(* IEC 61131-3 sources: PortalRobot/Portal_robot/Device/application/FB/FB_CELL_MANAGER, 14 files *)

(* ---- FB_CELL_MANAGER.st ---- *)
FUNCTION_BLOCK FB_CELL_MANAGER
VAR_INPUT
	xIoManual : BOOL; // Прямой ручной слой отменяет задание, не сбрасывая аварии
	axMagazineAutoSwapPending : ARRAY [1..GVL_CELL_SETTINGS.MagazineCount] OF BOOL; // Палета ждёт окна обмена
	axMagazineExchangeInProgress : ARRAY [1..GVL_CELL_SETTINGS.MagazineCount] OF BOOL; // Во время смены палет запрещены операции только с этим магазином
	xMagazineExchangeActive : BOOL; // Есть активный обмен палет; подавляет временные предупреждения о запасах
	xStart            : BOOL; // Импульс запуска цикла или отмены остановки
	xStop             : BOOL; // Импульс контролируемой остановки
	xTestAbort        : BOOL; // Немедленная отмена только тестового прогона
	xResetRequest     : BOOL; // Необработанный запрос сброса от HMI
	xReset            : BOOL; // Общий сброс владельцев ошибок
	xOperatorChoice   : BOOL; // Импульс ответа активному предпусковому опросу
	xOperatorCancel   : BOOL; // Импульс отмены предпускового опроса
	uiOperatorChoice  : UINT; // Выбранное содержимое, тип продукции или станок
	xManual           : BOOL; // Ручной режим ячейки
	xIoDoRejected : BOOL;
    xIoEmergencyResetRejected : BOOL;
    xIoEmergencyStopActive : BOOL;
	xIoOverrideRejected : BOOL; // Отклонённая транзакция диагностики, эффект WARNING
	xSettingsRejected : BOOL; // Rejected or expired setting transaction
	uiModeRejectReason : UINT; // Одноцикловый отказ транзакции режима: 2 цикл, 3 Safety
	xGlobalError      : BOOL; // Глобальная ошибка ячейки
	xSafetyReady      : BOOL; // Все дискретные условия безопасности выполнены
	xDrivesReady      : BOOL; // Приводы готовы
	xMotionBusy       : BOOL; // Оси ещё движутся
	xRobotInterfaceReady : BOOL; // Выбранный интерфейс робота готов к работе
	lrRobotActualX    : LREAL; // Фактическая координата робота X
	lrRobotActualY    : LREAL; // Фактическая координата робота Y
	lrRobotActualZ    : LREAL; // Фактическая координата робота Z
	stSafetyHomePoint : ST_POINT; // Настроенная безопасная точка повторного запуска
	lrSafetyHomeToleranceX : LREAL; // Допуск HOME_SAFETY по X
	lrSafetyHomeToleranceY : LREAL; // Допуск HOME_SAFETY по Y
	lrSafetyHomeToleranceZ : LREAL; // Допуск HOME_SAFETY по Z
	lrStoppedPoseTolerance : LREAL; // Допуск контроля позы после штатной остановки
	Config            : ST_MULTI_TYPE_CONFIG; // Активная конфигурация типов
	xConfigurationValid : BOOL; // Конфигурация типов прошла проверку
	xPointsConfigured : BOOL; // HOME_SAFETY и точки включённого оборудования настроены
	stRobotStatus     : ST_ROBOT_STATUS; // Состояние робота
	astMagazineStatus : ARRAY [1..GVL_CELL_SETTINGS.MagazineCount] OF ST_MAGAZINE_STATUS;
	astMachineStatus  : ARRAY [1..3] OF ST_MACHINE_PUBLIC; // Состояния станков
	astMachineDiag    : ARRAY [1..3] OF ST_MACHINE_DIAG; // Автоматы станков
	FaultRequest      : ST_CELL_FAULT_REQUEST; // Диагностическая инъекция
END_VAR
VAR_OUTPUT
	Command            : ST_CELL_COMMAND; // Команды существующим блокам ячейки
	Status             : ST_CELL_STATUS; // Общий контракт состояния ячейки
	Diag               : ST_CELL_DIAG; // Общий контракт диагностики ячейки
	Error              : ST_CELL_ERRORS; // Общий контракт ошибок ячейки
	CycleStatus        : ST_CELL_CYCLE_STATUS; // Расширенная диагностика универсального цикла
	FaultStatus        : ST_FAULT_INJECTION_STATUS; // Инъекция логической ошибки ячейки
	uiReturnMagazine   : UINT; // Внутренний владелец парного цикла до возврата детали; 0 — цикл освобождён
END_VAR
VAR
	axGeometryUnloadBlocked : ARRAY [1..3] OF BOOL; // Вызванная деталь ждёт доступного свободного ГК
	atonGeometryWait : ARRAY [1..3] OF TON;
	audiGeometryWaitCallId : ARRAY [1..3] OF UDINT;
	axGeometryWaitWarned : ARRAY [1..3] OF BOOL;
	xGeometryHeld : BOOL;
	xGeometryDetailCounted : BOOL;
	uiGeometryMachine : UINT;
	uiGeometryStation : UINT;
	uiGeometryParkStation : UINT;
	uiGeometryStep : UINT;
	uiGeometryBypassReason : UINT;
	uiGeometryIndex : UINT;
	udiGeometryMagazineCounter : UDINT;
	eGeometryReturnState : E_CELL_MANAGER_STATE;
	eGeometrySafePoint : E_POINT_NAME;
	eGeometryChangePoint : E_POINT_NAME;
	eGeometryPlacePoint : E_POINT_NAME;
	xActiveMagazineAutoSwapPending : BOOL; // Удержать владельца и цикл до обмена его палеты
	eState               : E_CELL_MANAGER_STATE := E_CELL_MANAGER_STATE.IDLE; // Состояние универсального автомата
	eMagazineOperation   : E_MAGAZINE_OPERATION; // Выполняемая операция магазина
	eMachineOperation    : E_MACHINE_OPERATION; // Зафиксированная операция станка
	xRunning             : BOOL; // Защёлка автоматического цикла
	xStopRequested       : BOOL; // Остановка после безопасного шага
	xReadyToStart        : BOOL; // Условия запуска выполнены
	xRobotReady          : BOOL; // Робот готов принять маршрут
	xMagazineReady       : BOOL; // Магазин готов к операции
	xActiveMagazineExchangeInProgress : BOOL; // Выбранный магазин сейчас меняет палеты
	stMagazineStatus     : ST_MAGAZINE_STATUS; // Снимок выбранного магазина для существующего автомата
	uiActiveMagazine     : UINT; // Магазин текущей команды роботу
	uiSupplyMagazine     : UINT; // Источник следующих заготовок сохраняется между парными циклами
	xMagazine1Available  : BOOL;
	xMagazine2Available  : BOOL;
	xMagazineSelectionAllowed : BOOL; // Новое владение допускается только между операциями
	xMagazine1CanContinue : BOOL; // Первый магазин позволяет следующий технологический шаг
	xMagazine2CanContinue : BOOL; // Второй магазин позволяет следующий технологический шаг
	xMagazine1CanSupplyBlank : BOOL; // М1 позволяет штатный план TAKE перед отдельной выгрузкой
	xMagazine2CanSupplyBlank : BOOL; // М2 позволяет штатный план TAKE перед отдельной выгрузкой
	xMagazine1CanExchangeDetail : BOOL; // Заготовка М1 освобождает слот для детали робота
	xMagazine2CanExchangeDetail : BOOL;
	xMagazine1CanPutDetail : BOOL; // Готовый магазин со свободным местом для детали робота
	xMagazine2CanPutDetail : BOOL;
	xActiveMagazineCanExchangeDetail : BOOL;
	xHeldBlankLoadAvailable : BOOL; // При двух грузах можно сначала загрузить пустой станок
	uiMagazineType       : UINT; // Тип станка при проверке содержимого обоих магазинов
	uiPreferredMagazine  : UINT; // Назначение с учётом владельца цикла и сохранённого источника
	xReselectMagazine    : BOOL; // Требуется передать владение подходящему магазину
	xAlternateMagazineAvailable : BOOL; // Второй магазин готов принять непрерывный автоматический цикл
	xUseAlternateMagazineForDetail : BOOL; // У текущего магазина нет слота детали, у второго есть
	xAnyMagazineDetailSlotAvailable : BOOL; // Есть доступный слот детали хотя бы в одном магазине
	xNoDetailDestinationCondition : BOOL; // Робот держит готовую деталь без доступного слота
	xNoBlankStockCondition : BOOL; // Нет заготовок и текущей работы для автоматического цикла
	xDetailDestinationWarningActive : BOOL; // Предупреждение об отсутствии места уже выдано
	xBlankStockWarningActive : BOOL; // Предупреждение об отсутствии заготовок уже выдано
	xMachineWorkPending : BOOL; // Станок занят/обрабатывает, запускается или содержит изделие
	xAnyMachineBusy      : BOOL; // Хотя бы один станок обслуживается
	xMachineServiceStarted : BOOL; // Выбранный станок вошёл в рецепт
	xReselectAfterRobotRelease : BOOL; // После снятия команды требуется повторный выбор
	xChangePrepared      : BOOL; // Для CHANGE зафиксированы совместимый станок и два корректных слота
	xFaultAllowed        : BOOL; // Инъекция разрешена в полностью остановленной ячейке
	xResetAllowed        : BOOL; // Локальная ошибка может быть сброшена
	xPayloadRouteWarningActive : BOOL; // Предупреждение о несовпадении типа груза и назначения уже выдано
	xPrestartGripper1Occupied : BOOL; // Снимок занятости первого захвата на момент запуска опроса
	xPrestartGripper2Occupied : BOOL; // Снимок занятости второго захвата на момент запуска опроса
	xSafetyHomeRequired : BOOL; // Защёлка обязательного возврата в HOME_SAFETY
	xRobotAtSafetyHome  : BOOL; // Робот находится в допустимом диапазоне HOME_SAFETY
	xStoppedPoseValid   : BOOL; // После штатной остановки сохранена доверенная поза
	xWasRunning         : BOOL; // Состояние цикла на предыдущем вызове
	xStartCheckCellIdle           : BOOL; // Отдельные условия запуска для HMI
	xStartCheckAutomaticMode      : BOOL;
	xStartCheckNoBlockingError    : BOOL;
	xStartCheckRobotInterfaceReady: BOOL;
	xStartCheckConfigurationValid : BOOL;
	xStartCheckPointsConfigured   : BOOL;
	xStartCheckDrivesReady        : BOOL;
	xStartCheckRobotReady         : BOOL;
	xStartCheckMagazineReady      : BOOL;
	xStartCheckTaskAvailable      : BOOL;
	xStartCheckSafetyHome         : BOOL;
	xStartCheckSafety             : BOOL;
	xOperatorPromptState          : BOOL; // Текущий шаг ожидает ответ HMI
	xOperatorChoiceAllowed        : BOOL;
	xOperatorCancelAllowed        : BOOL;
	uiOperatorPrompt              : UINT;
	uiOperatorTypeMask            : UINT;
	uiOperatorMachineMask         : UINT;
	uiStartConditionsMet         : UINT;
	lrStoppedPoseX      : LREAL; // Доверенная координата X штатной остановки
	lrStoppedPoseY      : LREAL; // Доверенная координата Y штатной остановки
	lrStoppedPoseZ      : LREAL; // Доверенная координата Z штатной остановки
	uiReadyMachines      : UINT; // Число доступных маршрутных целей
	uiMachine            : UINT; // Индекс станка
	uiMagazineIndex      : UINT; // Индекс магазина при поиске свободного слота
	uiCandidateMachine   : UINT; // Результат выбора
	uiSelectedMachine    : UINT; // Зафиксированный станок
	uiSelectedType       : UINT; // Тип маршрута
	uiBlankPayloadType   : UINT; // Тип заготовки в первом захвате
	uiDetailPayloadType  : UINT; // Тип готовой детали во втором захвате
	axMachineStartPending: ARRAY [1..3] OF BOOL; // Станок обслужен, но xProcessing ещё не подтверждён
	iTakeSlot            : SINT; // Зарезервированный слот заготовки
	iPutSlot             : SINT; // Зарезервированный слот укладки
	iTakeOriginSlot      : SINT; // Исходный слот заготовки для приоритетного возврата
	rtStart              : R_TRIG; // Фронт запуска
	rtStop               : R_TRIG; // Фронт остановки
	rtReset              : R_TRIG; // Фронт сброса
	rtOperatorChoice     : R_TRIG; // Один ответ не переносится на следующий шаг опроса
	rtOperatorCancel     : R_TRIG; // Фронт отмены предпускового опроса
	fbFaultInjector      : FB_CELL_FAULT_INJECTOR; // Проверка противоречивого груза
END_VAR
VAR CONSTANT
	FIRST_MACHINE     : UINT := UINT#1;
	LAST_MACHINE      : UINT := UINT#3;
	MACHINE_SWITCH_DEADBAND : TIME := T#1S; // Минимальный выигрыш времени для смены ожидаемой цели
	START_PENDING_ESTIMATE  : TIME := T#1S; // Оценка перехода от освобождения робота до xProcessing
	ERR_BOTH_GRIPPERS : DWORD := DWORD#16#0000_0001;
	ERR_ROBOT         : DWORD := DWORD#16#0000_0002;
	ERR_MAGAZINE      : DWORD := DWORD#16#0000_0004;
	ERR_MACHINE       : DWORD := DWORD#16#0000_0008;
	ERR_GLOBAL_STOP   : DWORD := DWORD#16#0000_0010;
	WRN_START_NOT_READY       : UINT := UINT#4;
	WRN_STOP_NOT_RUNNING      : UINT := UINT#5;
	WRN_SIM_ERROR_NOT_ALLOWED : UINT := UINT#8;
	WRN_PAYLOAD_ROUTE_MISMATCH : UINT := UINT#9;
	WRN_SAFETY_HOME_REQUIRED   : UINT := UINT#10;
	WRN_MANUAL_MODE_REJECTED   : UINT := UINT#11;
	WRN_CELL_SETTING_REJECTED : UINT := UINT#28;
	WRN_AUTOMATIC_MODE_REJECTED : UINT := UINT#27; // WARNING: общая авария удерживает ручной режим
	WRN_GRIPPER1_CONTENT       : UINT := UINT#15;
	WRN_GRIPPER2_CONTENT       : UINT := UINT#16;
	WRN_PAYLOAD_TYPE_CHOICE    : UINT := UINT#17;
	WRN_DETAIL_SLOT_REQUIRED   : UINT := UINT#18;
	WRN_START_MACHINE_REQUIRED : UINT := UINT#19;
	WRN_START_MACHINE_CHOICE   : UINT := UINT#20;
	WRN_OPERATOR_REPLY_REJECTED: UINT := UINT#21;
	WRN_OPERATOR_CANCEL_REJECTED: UINT := UINT#22;
	WRN_NO_DETAIL_DESTINATION  : UINT := UINT#29;
	WRN_NO_BLANK_STOCK         : UINT := UINT#30;
	WRN_GEOMETRY_WAIT_TIMEOUT  : UINT := UINT#52;
	WRN_IO_OVERRIDE_REJECTED   : UINT := UINT#31;
    WRN_IO_DO_REJECTED : UINT := UINT#32;
    WRN_IO_EMERGENCY_RESET_REJECTED : UINT := UINT#33;
END_VAR

// --- BEGIN IMPLEMENTATION ---

IF xIoDoRejected THEN
    Diag.stWarning.uiCode := WRN_IO_DO_REJECTED; // WARNING: вход/команда прямого ручного I/O не применены
    Diag.stWarning.udiSequence := Diag.stWarning.udiSequence + UDINT#1;
    IF Diag.stWarning.udiSequence = UDINT#0 THEN Diag.stWarning.udiSequence := UDINT#1; END_IF;
END_IF;
IF xIoEmergencyResetRejected THEN
    Diag.stWarning.uiCode := WRN_IO_EMERGENCY_RESET_REJECTED; // WARNING: останов остаётся
    Diag.stWarning.udiSequence := Diag.stWarning.udiSequence + UDINT#1;
    IF Diag.stWarning.udiSequence = UDINT#0 THEN Diag.stWarning.udiSequence := UDINT#1; END_IF;
END_IF;
IF xIoOverrideRejected THEN
    Diag.stWarning.uiCode := WRN_IO_OVERRIDE_REJECTED; // WARNING: входы не изменены
    Diag.stWarning.udiSequence := Diag.stWarning.udiSequence + UDINT#1;
    IF Diag.stWarning.udiSequence = UDINT#0 THEN Diag.stWarning.udiSequence := UDINT#1; END_IF;
END_IF;
IF xSettingsRejected THEN
	Diag.stWarning.uiCode := WRN_CELL_SETTING_REJECTED; // WARNING: settings unchanged
	Diag.stWarning.udiSequence := Diag.stWarning.udiSequence + UDINT#1;
	IF Diag.stWarning.udiSequence = UDINT#0 THEN Diag.stWarning.udiSequence := UDINT#1; END_IF;
END_IF;

rtStart(CLK := xStart);
rtStop(CLK := xStop);
rtReset(CLK := xResetRequest);
rtOperatorChoice(CLK := xOperatorChoice);
rtOperatorCancel(CLK := xOperatorCancel);

// До выбора магазина/станка исключаем выгрузку вызванной детали без свободного ГК.
UpdateGeometryWait();

// Выбор выполняется только между операциями. Внутренний автомат по-прежнему
// работает с одним снимком, поэтому уже отлажанный маршрут не размазывается
// по двум владельцам и не переключается посреди TAKE/CHANGE.
xMagazine1Available := astMagazineStatus[1].xEnabled
	AND astMagazineStatus[1].xReady
	AND NOT axMagazineAutoSwapPending[1]
	AND NOT axMagazineExchangeInProgress[1]
	AND NOT astMagazineStatus[1].xBusy
	AND NOT astMagazineStatus[1].xError
	AND NOT astMagazineStatus[1].xDisablePending
	AND NOT astMagazineStatus[1].xFinished;
xMagazine2Available := astMagazineStatus[2].xEnabled
	AND astMagazineStatus[2].xReady
	AND NOT axMagazineAutoSwapPending[2]
	AND NOT axMagazineExchangeInProgress[2]
	AND NOT astMagazineStatus[2].xBusy
	AND NOT astMagazineStatus[2].xError
	AND NOT astMagazineStatus[2].xDisablePending
	AND NOT astMagazineStatus[2].xFinished;

// Реальная свободная позиция имеет приоритет перед дополнительным TAKE ради
// освобождения места. Индекс типа проверяется до чтения массивов.
xMagazine1CanPutDetail := FALSE;
xMagazine2CanPutDetail := FALSE;
IF stRobotStatus.xDetailAvailable
AND (uiDetailPayloadType >= UINT#1)
AND (uiDetailPayloadType <= Config.uiTypeCount)
AND (uiDetailPayloadType <= UINT#3) THEN
	xMagazine1CanPutDetail := xMagazine1Available
		AND (astMagazineStatus[1].stTypeStatus.aiFreeSlot[uiDetailPayloadType] > SINT#0);
	xMagazine2CanPutDetail := xMagazine2Available
		AND (astMagazineStatus[2].stTypeStatus.aiFreeSlot[uiDetailPayloadType] > SINT#0);
END_IF;

// Полная палета тоже принимает деталь: сначала берём заготовку свободным
// захватом 1, затем кладём деталь в освободившийся универсальный слот.
// Заготовке нужен совместимый маршрут; станок может ещё обрабатывать изделие.
xMagazine1CanExchangeDetail := FALSE;
xMagazine2CanExchangeDetail := FALSE;
xHeldBlankLoadAvailable := FALSE;
FOR uiMachine := FIRST_MACHINE TO LAST_MACHINE DO
	IF IsMachineEligible(uiMachine := uiMachine) THEN
		uiMagazineType := Config.auiMachineType[uiMachine];
		IF stRobotStatus.xBlankAvailable AND stRobotStatus.xDetailAvailable
		AND (uiMagazineType = uiBlankPayloadType)
		AND astMachineStatus[uiMachine].xCanAcceptService
		AND (astMachineStatus[uiMachine].ePartState = E_PART_STATE.EMPTY) THEN
			xHeldBlankLoadAvailable := TRUE;
		END_IF;
		IF stRobotStatus.xDetailAvailable
		AND NOT stRobotStatus.xBlankAvailable
		AND stRobotStatus.xGripper1Open
		AND (uiDetailPayloadType >= UINT#1)
		AND (uiDetailPayloadType <= Config.uiTypeCount)
		AND (uiMagazineType >= UINT#1) AND (uiMagazineType <= UINT#3)
		AND (astMachineStatus[uiMachine].xProcessing
			OR axMachineStartPending[uiMachine]
			OR (astMachineStatus[uiMachine].xCanAcceptService
				AND ((astMachineStatus[uiMachine].ePartState = E_PART_STATE.EMPTY)
					OR astMachineStatus[uiMachine].xServiceRequired))) THEN
			IF astMagazineStatus[1].stTypeStatus.aiBlankSlot[uiMagazineType] > SINT#0 THEN
				xMagazine1CanExchangeDetail := xMagazine1Available
					AND ((uiReturnMagazine = UINT#0) OR (uiReturnMagazine = UINT#1));
			END_IF;
			IF astMagazineStatus[2].stTypeStatus.aiBlankSlot[uiMagazineType] > SINT#0 THEN
				xMagazine2CanExchangeDetail := xMagazine2Available
					AND ((uiReturnMagazine = UINT#0) OR (uiReturnMagazine = UINT#2));
			END_IF;
		END_IF;
	END_IF;
END_FOR;

// После полной выработки или операторского запроса отключения активного магазина
// автомат не требует нового Start. Переключение выполняется только когда робот
// и старый магазин уже освобождены.
xAlternateMagazineAvailable := FALSE;
IF uiActiveMagazine = UINT#1 THEN
	xAlternateMagazineAvailable := xMagazine2Available;
ELSIF uiActiveMagazine = UINT#2 THEN
	xAlternateMagazineAvailable := xMagazine1Available;
END_IF;

// Если деталь уже у робота, сначала переключаем владение на второй магазин,
// если там есть совместимый свободный слот. Это происходит только на границе
// операций и не прерывает уже выданную команду.
xUseAlternateMagazineForDetail := FALSE;
IF xRunning
AND stRobotStatus.xDetailAvailable
AND ((eState = E_CELL_MANAGER_STATE.PLAN_TARGET)
	OR (eState = E_CELL_MANAGER_STATE.WAIT_TARGET)
	OR (eState = E_CELL_MANAGER_STATE.SELECT_FALLBACK)
	OR (eState = E_CELL_MANAGER_STATE.WAIT_MAGAZINE))
AND (uiDetailPayloadType >= UINT#1)
AND (uiDetailPayloadType <= Config.uiTypeCount) THEN
	IF uiActiveMagazine = UINT#1 THEN
		xUseAlternateMagazineForDetail := NOT xMagazine1CanPutDetail AND xMagazine2CanPutDetail;
	ELSIF uiActiveMagazine = UINT#2 THEN
		xUseAlternateMagazineForDetail := NOT xMagazine2CanPutDetail AND xMagazine1CanPutDetail;
	END_IF;
END_IF;
// На каждой границе планирования проверяем ОБА магазина. Готовность механики
// сама по себе не означает наличие следующей операции: учитываем типы заготовок
// и возможность вернуть изделие из включённого исправного станка.
// Уже взятую заготовку сначала обслуживаем или возвращаем в исходный слот.
xMagazineSelectionAllowed := NOT stRobotStatus.xBusy
	AND NOT stRobotStatus.xBlankAvailable
	AND ((eState = E_CELL_MANAGER_STATE.IDLE)
		OR (eState = E_CELL_MANAGER_STATE.PLAN_TARGET)
		OR (eState = E_CELL_MANAGER_STATE.WAIT_TARGET)
		OR (eState = E_CELL_MANAGER_STATE.SELECT_FALLBACK)
		OR (eState = E_CELL_MANAGER_STATE.WAIT_MAGAZINE));
xMagazine1CanContinue := xMagazine1Available;
xMagazine2CanContinue := xMagazine2Available;
xMagazine1CanSupplyBlank := FALSE;
xMagazine2CanSupplyBlank := FALSE;
IF xMagazineSelectionAllowed THEN
	xMagazine1CanContinue := FALSE;
	xMagazine2CanContinue := FALSE;
	IF stRobotStatus.xDetailAvailable THEN
		IF (uiDetailPayloadType >= UINT#1)
		AND (uiDetailPayloadType <= Config.uiTypeCount)
		AND (uiDetailPayloadType <= UINT#3) THEN
			xMagazine1CanContinue := xMagazine1Available
				AND ((astMagazineStatus[1].stTypeStatus.aiFreeSlot[uiDetailPayloadType] > SINT#0)
					OR xMagazine1CanExchangeDetail);
			xMagazine2CanContinue := xMagazine2Available
				AND ((astMagazineStatus[2].stTypeStatus.aiFreeSlot[uiDetailPayloadType] > SINT#0)
					OR xMagazine2CanExchangeDetail);
		END_IF;
	ELSE
		xMagazine1CanSupplyBlank := xMagazine1Available
			AND HasMagazineWork(uiMagazine := UINT#1, xSupplyBlankOnly := TRUE);
		xMagazine2CanSupplyBlank := xMagazine2Available
			AND HasMagazineWork(uiMagazine := UINT#2, xSupplyBlankOnly := TRUE);
		xMagazine1CanContinue := xMagazine1Available
			AND HasMagazineWork(uiMagazine := UINT#1, xSupplyBlankOnly := FALSE);
		xMagazine2CanContinue := xMagazine2Available
			AND HasMagazineWork(uiMagazine := UINT#2, xSupplyBlankOnly := FALSE);
	END_IF;
END_IF;
// PUT возвращается в магазин взятой заготовки. Резервная укладка не меняет источник.
// Между циклами дорабатываем выбранную палету; М1 имеет приоритет при первом выборе.
uiPreferredMagazine := UINT#0;
IF xMagazine1CanPutDetail AND (uiReturnMagazine = UINT#1) THEN
	uiPreferredMagazine := UINT#1;
ELSIF xMagazine2CanPutDetail AND (uiReturnMagazine = UINT#2) THEN
	uiPreferredMagazine := UINT#2;
ELSIF xMagazine1CanPutDetail THEN
	uiPreferredMagazine := UINT#1;
ELSIF xMagazine2CanPutDetail THEN
	uiPreferredMagazine := UINT#2;
ELSIF stRobotStatus.xDetailAvailable AND xMagazine1CanContinue
AND (uiReturnMagazine = UINT#1) THEN
	uiPreferredMagazine := UINT#1;
ELSIF stRobotStatus.xDetailAvailable AND xMagazine2CanContinue
AND (uiReturnMagazine = UINT#2) THEN
	uiPreferredMagazine := UINT#2;
ELSIF (uiSupplyMagazine = UINT#1) AND xMagazine1CanSupplyBlank THEN
	uiPreferredMagazine := UINT#1;
ELSIF (uiSupplyMagazine = UINT#2) AND xMagazine2CanSupplyBlank THEN
	uiPreferredMagazine := UINT#2;
ELSIF xMagazine1CanSupplyBlank THEN
	uiPreferredMagazine := UINT#1;
ELSIF xMagazine2CanSupplyBlank THEN
	uiPreferredMagazine := UINT#2;
ELSIF (uiSupplyMagazine = UINT#1) AND xMagazine1CanContinue THEN
	uiPreferredMagazine := UINT#1;
ELSIF (uiSupplyMagazine = UINT#2) AND xMagazine2CanContinue THEN
	uiPreferredMagazine := UINT#2;
ELSIF xMagazine1CanContinue THEN
	uiPreferredMagazine := UINT#1;
ELSIF xMagazine2CanContinue THEN
	uiPreferredMagazine := UINT#2;
END_IF;
xReselectMagazine := xMagazineSelectionAllowed
	AND (uiPreferredMagazine > UINT#0)
	AND (uiActiveMagazine <> uiPreferredMagazine)
	AND NOT ((uiActiveMagazine = UINT#1) AND astMagazineStatus[1].xBusy)
	AND NOT ((uiActiveMagazine = UINT#2) AND astMagazineStatus[2].xBusy);

IF xRunning
AND (eState <> E_CELL_MANAGER_STATE.GEOMETRY_WAIT_FREE)
AND (eState <> E_CELL_MANAGER_STATE.GEOMETRY_DELIVER)
AND (eState <> E_CELL_MANAGER_STATE.GEOMETRY_RELEASE_COMMAND)
AND (uiActiveMagazine >= UINT#1)
AND (uiActiveMagazine <= UINT#2) THEN
	// Операторское отключение активного магазина передаёт владение второму
	// только на границе операций. Фактический груз FB_ROBOT при этом остаётся
	// источником истины и будет уложен уже в выбранный магазин. Проверяем также
	// итоговый xEnabled: FB_MAGAZINE может завершить отключение и снять
	// xDisablePending раньше, чем робот достигнет границы перепланирования.
	// xFinished в DONE ещё не означает конец цикла: до завершения RELEASE_MAGAZINE
	// не меняем владельца. Когда началась сама смена палет, адресная блокировка
	// снимает старого владельца на границе операций и разрешает выбрать второй магазин.
	IF (((astMagazineStatus[uiActiveMagazine].xFinished
			AND NOT axMagazineAutoSwapPending[uiActiveMagazine])
		OR ((astMagazineStatus[uiActiveMagazine].xDisablePending
			OR NOT astMagazineStatus[uiActiveMagazine].xEnabled)
			AND ((eState = E_CELL_MANAGER_STATE.PLAN_TARGET)
				OR (eState = E_CELL_MANAGER_STATE.WAIT_TARGET)
				OR (eState = E_CELL_MANAGER_STATE.SELECT_FALLBACK)
				OR (eState = E_CELL_MANAGER_STATE.WAIT_MAGAZINE))))
		OR axMagazineExchangeInProgress[uiActiveMagazine]
		OR xUseAlternateMagazineForDetail
		OR xReselectMagazine)
	AND (NOT astMagazineStatus[uiActiveMagazine].xBusy
		OR axMagazineExchangeInProgress[uiActiveMagazine])
	AND NOT stRobotStatus.xBusy THEN
		IF xAlternateMagazineAvailable THEN
			IF uiActiveMagazine = UINT#1 THEN
				uiActiveMagazine := UINT#2;
			ELSE
				uiActiveMagazine := UINT#1;
			END_IF;
		ELSE
			// Без готовой замены старый код навечно оставлял магазин владельцем:
			// FB_MAGAZINE видел xRobotOwnsMagazine и не мог завершить Disable.
			// Освобождаем владение и ждём готовый магазин, не останавливая ячейку.
			uiActiveMagazine := UINT#0;
		END_IF;
		eMagazineOperation := E_MAGAZINE_OPERATION.NONE;
		eMachineOperation := E_MACHINE_OPERATION.NONE;
		uiSelectedMachine := UINT#0;
		uiSelectedType := UINT#0;
		iTakeSlot := SINT#0;
		iPutSlot := SINT#0;
		iTakeOriginSlot := SINT#0;
		IF uiActiveMagazine = UINT#0 THEN
			eState := E_CELL_MANAGER_STATE.WAIT_MAGAZINE;
		ELSE
			eState := E_CELL_MANAGER_STATE.PLAN_TARGET;
		END_IF;
	END_IF;
END_IF;

IF (uiActiveMagazine < UINT#1) OR (uiActiveMagazine > UINT#2) THEN
	IF uiPreferredMagazine > UINT#0 THEN
		uiActiveMagazine := uiPreferredMagazine;
	ELSIF xMagazine1Available THEN
		uiActiveMagazine := UINT#1;
	ELSIF xMagazine2Available THEN
		uiActiveMagazine := UINT#2;
	ELSE
		uiActiveMagazine := UINT#0;
	END_IF;
ELSIF NOT xRunning
AND (astMagazineStatus[uiActiveMagazine].xFinished
	OR astMagazineStatus[uiActiveMagazine].xError
	OR NOT astMagazineStatus[uiActiveMagazine].xEnabled
	OR xReselectMagazine) THEN
	IF (uiActiveMagazine <> UINT#1) AND xMagazine1Available THEN
		uiActiveMagazine := UINT#1;
	ELSIF (uiActiveMagazine <> UINT#2) AND xMagazine2Available THEN
		uiActiveMagazine := UINT#2;
	ELSIF xMagazine1Available THEN
		uiActiveMagazine := UINT#1;
	ELSIF xMagazine2Available THEN
		uiActiveMagazine := UINT#2;
	ELSE
		uiActiveMagazine := UINT#0;
	END_IF;
END_IF;

xActiveMagazineCanExchangeDetail := ((uiActiveMagazine = UINT#1) AND xMagazine1CanExchangeDetail)
	OR ((uiActiveMagazine = UINT#2) AND xMagazine2CanExchangeDetail);

IF (uiActiveMagazine >= UINT#1) AND (uiActiveMagazine <= UINT#2) THEN
	stMagazineStatus := astMagazineStatus[uiActiveMagazine];
	xActiveMagazineAutoSwapPending := axMagazineAutoSwapPending[uiActiveMagazine];
	xActiveMagazineExchangeInProgress := axMagazineExchangeInProgress[uiActiveMagazine];
ELSE
	stMagazineStatus := astMagazineStatus[1];
	xActiveMagazineAutoSwapPending := FALSE;
	xActiveMagazineExchangeInProgress := axMagazineExchangeInProgress[1];
END_IF;

// HOME_SAFETY — это диапазон вокруг именованной точки, а не требование
// побитового совпадения координат. Защёлка снимается только при принятом запуске:
// оператор не сможет подъехать к точке, снова отъехать и запустить цикл.
xRobotAtSafetyHome := (ABS(lrRobotActualX - stSafetyHomePoint.X) <= lrSafetyHomeToleranceX)
	AND (ABS(lrRobotActualY - stSafetyHomePoint.Y) <= lrSafetyHomeToleranceY)
	AND (ABS(lrRobotActualZ - stSafetyHomePoint.Z) <= lrSafetyHomeToleranceZ);

// Штатная остановка не требует HOME_SAFETY, пока робот остаётся в сохранённой
// позе. Любое последующее координатное перемещение (JOG, MoveAbsolute или
// MoveDirect) необратимо снимает доверие до следующего разрешённого запуска.
IF (eState = E_CELL_MANAGER_STATE.IDLE)
AND NOT xRunning
AND NOT xSafetyHomeRequired THEN
	IF NOT xStoppedPoseValid THEN
		lrStoppedPoseX := lrRobotActualX;
		lrStoppedPoseY := lrRobotActualY;
		lrStoppedPoseZ := lrRobotActualZ;
		xStoppedPoseValid := TRUE;
	ELSIF xManual
	AND ((ABS(lrRobotActualX - lrStoppedPoseX) > lrStoppedPoseTolerance)
	OR (ABS(lrRobotActualY - lrStoppedPoseY) > lrStoppedPoseTolerance)
	OR (ABS(lrRobotActualZ - lrStoppedPoseZ) > lrStoppedPoseTolerance)) THEN
		xSafetyHomeRequired := TRUE;
		xStoppedPoseValid := FALSE;
	END_IF;
END_IF;

// FB_ROBOT — источник фактического типа груза. Локальные значения менеджера
// принимаются от него после каждого цикла, что оставляет место для будущей
// инициализации зажатого захвата оператором.
IF stRobotStatus.xBlankAvailable THEN
	uiBlankPayloadType := stRobotStatus.uiBlankPayloadType;
ELSE
	uiBlankPayloadType := UINT#0;
END_IF;
IF stRobotStatus.xDetailAvailable THEN
	uiDetailPayloadType := stRobotStatus.uiDetailPayloadType;
ELSE
	uiDetailPayloadType := UINT#0;
END_IF;

// FB_MACHINE остаётся единственным владельцем таймаута запуска. Диспетчер только
// сохраняет короткое переходное состояние, чтобы новый цикл не исключался из прогноза.
FOR uiMachine := FIRST_MACHINE TO LAST_MACHINE DO
	IF axMachineStartPending[uiMachine]
	AND (astMachineStatus[uiMachine].xProcessing
		OR (astMachineStatus[uiMachine].ePartState = E_PART_STATE.EMPTY)
		OR NOT astMachineStatus[uiMachine].xEnabled
		OR astMachineStatus[uiMachine].xDisablePending
		OR astMachineStatus[uiMachine].xError) THEN
		axMachineStartPending[uiMachine] := FALSE;
	END_IF;
END_FOR;

Command.stRobot.xExecute := FALSE;
FOR uiGeometryIndex := UINT#1 TO UINT#2 DO
	GVL_GEOMETRY_CONTROL.astSignals[uiGeometryIndex].xReleased := FALSE;
END_FOR;
// После аварии контекст снимается лишь при подтверждённом выходе в HOME_SAFETY.
IF (uiGeometryStation >= UINT#1) AND (uiGeometryStation <= UINT#2)
AND (stRobotStatus.eCurrentPoint = E_POINT_NAME.HOME_SAFETY)
AND NOT stRobotStatus.xBusy AND NOT xMotionBusy
AND (eState <> E_CELL_MANAGER_STATE.GEOMETRY_DELIVER)
AND (eState <> E_CELL_MANAGER_STATE.GEOMETRY_RELEASE_COMMAND) THEN
	GVL_GEOMETRY_CONTROL.astSignals[uiGeometryStation].xReserve := FALSE;
	GVL_GEOMETRY_CONTROL.astSignals[uiGeometryStation].xDeposited := FALSE;
	GVL_GEOMETRY_CONTROL.astSignals[uiGeometryStation].xRobotInteraction := FALSE;
	GVL_GEOMETRY_CONTROL.astSignals[uiGeometryStation].xReleased := TRUE;
	IF xGeometryHeld AND (uiGeometryMachine >= UINT#1) AND (uiGeometryMachine <= UINT#3)
	AND stRobotStatus.xDetailAvailable THEN
		GVL_GEOMETRY_CONTROL.astCalls[uiGeometryMachine].uiStation := UINT#0;
		GVL_GEOMETRY_CONTROL.astCalls[uiGeometryMachine].uiState := UINT#2;
		GVL_GEOMETRY_CONTROL.astCalls[uiGeometryMachine].uiReason := UINT#4;
		F_GEOMETRY_EVENT(Call := GVL_GEOMETRY_CONTROL.astCalls[uiGeometryMachine]);
	END_IF;
	IF NOT stRobotStatus.xDetailAvailable THEN
		IF xGeometryHeld AND (uiGeometryMachine >= UINT#1) AND (uiGeometryMachine <= UINT#3) THEN
			IF (GVL_GEOMETRY_CONTROL.astCalls[uiGeometryMachine].uiState = UINT#2)
			OR (GVL_GEOMETRY_CONTROL.astCalls[uiGeometryMachine].uiState = UINT#3) THEN
				GVL_GEOMETRY_CONTROL.astCalls[uiGeometryMachine].uiState := UINT#7;
				GVL_GEOMETRY_CONTROL.astCalls[uiGeometryMachine].uiReason := UINT#5;
				F_GEOMETRY_EVENT(Call := GVL_GEOMETRY_CONTROL.astCalls[uiGeometryMachine]);
			END_IF;
		END_IF;
		xGeometryHeld := FALSE; uiGeometryMachine := UINT#0;
	END_IF;
	uiGeometryStation := UINT#0;
END_IF;
// Ручное изъятие из захвата после остановки завершает старый вызов. Подтверждённую
// укладку на ГК (state 4) этот путь не заменяет прерыванием и повторно не считает.
IF xGeometryHeld AND NOT stRobotStatus.xDetailAvailable AND NOT xRunning
AND NOT stRobotStatus.xBusy AND NOT xMotionBusy
AND (eState = E_CELL_MANAGER_STATE.IDLE)
AND (uiGeometryMachine >= UINT#1) AND (uiGeometryMachine <= UINT#3) THEN
	IF (GVL_GEOMETRY_CONTROL.astCalls[uiGeometryMachine].uiState = UINT#2)
	OR (GVL_GEOMETRY_CONTROL.astCalls[uiGeometryMachine].uiState = UINT#3) THEN
		GVL_GEOMETRY_CONTROL.astCalls[uiGeometryMachine].uiState := UINT#7;
		GVL_GEOMETRY_CONTROL.astCalls[uiGeometryMachine].uiReason := UINT#5;
		F_GEOMETRY_EVENT(Call := GVL_GEOMETRY_CONTROL.astCalls[uiGeometryMachine]);
	END_IF;
	xGeometryHeld := FALSE; uiGeometryMachine := UINT#0;
END_IF;
Command.stRobot.xStop := FALSE;
Command.stRobot.xReset := xReset;
Command.stRobot.eAction := E_ROBOT_ACTION.NONE;
Command.stRobot.eSetPoint := E_POINT_NAME.NONE;
Command.stRobot.iActiveSlot := SINT#0;
Command.stRobot.uiMagazineId := UINT#0;
Command.uiBlankPayloadType := uiBlankPayloadType;
Command.uiDetailPayloadType := uiDetailPayloadType;

Command.stMagazine.xEnable := FALSE;
Command.stMagazine.xDisable := FALSE;
Command.stMagazine.xExecute := FALSE;
Command.stMagazine.xStop := FALSE;
Command.stMagazine.eOperation := eMagazineOperation;
Command.stMagazine.iTakeSlot := iTakeSlot;
Command.stMagazine.iPutSlot := iPutSlot;
xChangePrepared := FALSE;

FOR uiMachine := FIRST_MACHINE TO LAST_MACHINE DO
	Command.axMachineExecute[uiMachine] := FALSE;
END_FOR;

uiReadyMachines := UINT#0;
xAnyMachineBusy := FALSE;
xMachineWorkPending := FALSE;
FOR uiMachine := FIRST_MACHINE TO LAST_MACHINE DO
	IF astMachineStatus[uiMachine].xBusy THEN
		xAnyMachineBusy := TRUE;
		xMachineWorkPending := TRUE;
	END_IF;
	IF astMachineStatus[uiMachine].xProcessing
	OR astMachineStatus[uiMachine].xPartReady
	OR axMachineStartPending[uiMachine]
	OR ((astMachineStatus[uiMachine].ePartState = E_PART_STATE.LOADED)
		AND ((astMachineStatus[uiMachine].ePartType = E_PART_TYPE.PART)
			OR (astMachineStatus[uiMachine].ePartType = E_PART_TYPE.DETAIL))) THEN
		xMachineWorkPending := TRUE;
	END_IF;
	IF IsMachineEligible(uiMachine := uiMachine) THEN
		uiReadyMachines := uiReadyMachines + UINT#1;
	END_IF;
END_FOR;

xRobotReady := NOT stRobotStatus.xBusy
	AND NOT stRobotStatus.xError;
xMagazineReady := (uiActiveMagazine >= UINT#1)
	AND (uiActiveMagazine <= UINT#2)
	AND NOT xActiveMagazineExchangeInProgress
	AND NOT xActiveMagazineAutoSwapPending
	AND stMagazineStatus.xEnabled
	AND stMagazineStatus.xReady
	AND NOT stMagazineStatus.xBusy
	AND NOT stMagazineStatus.xError
	AND NOT stMagazineStatus.xFinished
	AND NOT stMagazineStatus.xDisablePending;

uiCandidateMachine := SelectMachineBeforeTake();
IF uiCandidateMachine = UINT#0 THEN
	uiCandidateMachine := SelectMachineForUnload(uiCurrentMachine := UINT#0);
END_IF;

// Для готовой детали пригоден только свободный слот её типа в магазине,
// который сейчас включён и доступен роботу. Свободная ячейка в отключённом
// или неисправном магазине не считается маршрутом.
xAnyMagazineDetailSlotAvailable := FALSE;
IF (uiDetailPayloadType >= UINT#1)
AND (uiDetailPayloadType <= Config.uiTypeCount) THEN
	FOR uiMagazineIndex := UINT#1 TO GVL_CELL_SETTINGS.MagazineCount DO
		IF astMagazineStatus[uiMagazineIndex].xEnabled
		AND astMagazineStatus[uiMagazineIndex].xReady
		AND NOT axMagazineExchangeInProgress[uiMagazineIndex]
		AND NOT axMagazineAutoSwapPending[uiMagazineIndex]
		AND NOT astMagazineStatus[uiMagazineIndex].xBusy
		AND NOT astMagazineStatus[uiMagazineIndex].xError
		AND NOT astMagazineStatus[uiMagazineIndex].xFinished
		AND NOT astMagazineStatus[uiMagazineIndex].xDisablePending THEN
			IF astMagazineStatus[uiMagazineIndex].stTypeStatus.aiFreeSlot[uiDetailPayloadType] > SINT#0 THEN
				xAnyMagazineDetailSlotAvailable := TRUE;
			END_IF;
		END_IF;
	END_FOR;
END_IF;

// WARNING: место требуется только для готовой детали, уже находящейся у робота.
// Деталь в станке и полная палета заготовок при пустом роботе не создают W29.
// Взятие заготовки освобождает место; при двух грузах возможна загрузка станка.
// Штатный Stop снимает потребность в новом маршруте. Фронт проверяем отдельно:
// защёлка xStopRequested обновляется ниже, после регистрации предупреждений.
xNoDetailDestinationCondition := (xRunning OR rtStart.Q)
	AND NOT rtStop.Q
	AND NOT xStopRequested
	AND NOT xManual
	AND NOT xMagazineExchangeActive
	AND stRobotStatus.xDetailAvailable
	AND (uiDetailPayloadType >= UINT#1)
	AND (uiDetailPayloadType <= Config.uiTypeCount)
	AND NOT xAnyMagazineDetailSlotAvailable
	AND NOT xMagazine1CanExchangeDetail
	AND NOT xMagazine2CanExchangeDetail
	AND NOT xHeldBlankLoadAvailable
	AND ((eState = E_CELL_MANAGER_STATE.PLAN_TARGET)
		OR (eState = E_CELL_MANAGER_STATE.WAIT_TARGET)
		OR (eState = E_CELL_MANAGER_STATE.SELECT_FALLBACK)
		OR (eState = E_CELL_MANAGER_STATE.WAIT_MAGAZINE)
		OR (rtStart.Q AND (eState = E_CELL_MANAGER_STATE.IDLE)));

xNoBlankStockCondition := (xRunning OR rtStart.Q)
	AND NOT xManual
	AND NOT xMagazineExchangeActive
	AND NOT stRobotStatus.xBlankAvailable
	AND NOT stRobotStatus.xDetailAvailable
	AND astMagazineStatus[1].xOutBlank
	AND astMagazineStatus[2].xOutBlank
	AND NOT xMachineWorkPending
	AND (uiCandidateMachine = UINT#0)
	AND ((eState = E_CELL_MANAGER_STATE.PLAN_TARGET)
		OR (eState = E_CELL_MANAGER_STATE.WAIT_TARGET)
		OR (eState = E_CELL_MANAGER_STATE.WAIT_MAGAZINE)
		OR (rtStart.Q AND (eState = E_CELL_MANAGER_STATE.IDLE)));

CASE Config.uiTypeCount OF
	UINT#1: uiOperatorTypeMask := UINT#1;
	UINT#2: uiOperatorTypeMask := UINT#3;
	UINT#3: uiOperatorTypeMask := UINT#7;
ELSE
	uiOperatorTypeMask := UINT#0;
END_CASE;

// Для специального старта с двумя грузами оператор выбирает только среди действительно
// пустых, готовых и совместимых станков. Окончательная проверка выбора остаётся в PLC.
uiOperatorMachineMask := UINT#0;
IF (uiBlankPayloadType >= UINT#1)
AND (uiBlankPayloadType <= Config.uiTypeCount) THEN
	FOR uiMachine := FIRST_MACHINE TO LAST_MACHINE DO
		IF IsMachineCompatible(
			uiMachine := uiMachine,
			uiProductType := uiBlankPayloadType
		)
		AND astMachineStatus[uiMachine].xCanAcceptService
		AND (astMachineStatus[uiMachine].ePartState = E_PART_STATE.EMPTY) THEN
			CASE uiMachine OF
				UINT#1: uiOperatorMachineMask := uiOperatorMachineMask OR UINT#1;
				UINT#2: uiOperatorMachineMask := uiOperatorMachineMask OR UINT#2;
				UINT#3: uiOperatorMachineMask := uiOperatorMachineMask OR UINT#4;
			END_CASE;
		END_IF;
	END_FOR;
END_IF;

// Условия запуска публикуются раздельно: PLC остаётся единственным владельцем
// технологического решения, а HMI только объясняет его оператору.
xStartCheckCellIdle := (eState = E_CELL_MANAGER_STATE.IDLE) AND NOT xRunning;
xStartCheckAutomaticMode := NOT xManual;
xStartCheckNoBlockingError := NOT xGlobalError AND NOT xIoManual AND (Error.dwErrorActive = DWORD#0);
xStartCheckRobotInterfaceReady := xRobotInterfaceReady;
xStartCheckConfigurationValid := xConfigurationValid;
xStartCheckPointsConfigured := xPointsConfigured;
xStartCheckDrivesReady := xDrivesReady;
xStartCheckRobotReady := xRobotReady;
xStartCheckMagazineReady := xMagazineReady;
xStartCheckTaskAvailable := stRobotStatus.xBlankAvailable
		OR stRobotStatus.xDetailAvailable
		OR (uiCandidateMachine > UINT#0);
xStartCheckSafetyHome := NOT xSafetyHomeRequired OR xRobotAtSafetyHome;
xStartCheckSafety := xSafetyReady;

xReadyToStart := xStartCheckCellIdle
	AND xStartCheckAutomaticMode
	AND xStartCheckNoBlockingError
	AND xStartCheckRobotInterfaceReady
	AND xStartCheckConfigurationValid
	AND xStartCheckPointsConfigured
	AND xStartCheckDrivesReady
	AND xStartCheckRobotReady
	AND xStartCheckMagazineReady
	AND xStartCheckTaskAvailable
	AND xStartCheckSafetyHome
	AND xStartCheckSafety;

uiStartConditionsMet := UINT#0;
IF xStartCheckCellIdle THEN
	uiStartConditionsMet := uiStartConditionsMet + UINT#1;
END_IF;
IF xStartCheckAutomaticMode THEN
	uiStartConditionsMet := uiStartConditionsMet + UINT#1;
END_IF;
IF xStartCheckNoBlockingError THEN
	uiStartConditionsMet := uiStartConditionsMet + UINT#1;
END_IF;
IF xStartCheckRobotInterfaceReady THEN
	uiStartConditionsMet := uiStartConditionsMet + UINT#1;
END_IF;
IF xStartCheckConfigurationValid THEN
	uiStartConditionsMet := uiStartConditionsMet + UINT#1;
END_IF;
IF xStartCheckPointsConfigured THEN
	uiStartConditionsMet := uiStartConditionsMet + UINT#1;
END_IF;
IF xStartCheckDrivesReady THEN
	uiStartConditionsMet := uiStartConditionsMet + UINT#1;
END_IF;
IF xStartCheckRobotReady THEN
	uiStartConditionsMet := uiStartConditionsMet + UINT#1;
END_IF;
IF xStartCheckMagazineReady THEN
	uiStartConditionsMet := uiStartConditionsMet + UINT#1;
END_IF;
IF xStartCheckTaskAvailable THEN
	uiStartConditionsMet := uiStartConditionsMet + UINT#1;
END_IF;
IF xStartCheckSafetyHome THEN
	uiStartConditionsMet := uiStartConditionsMet + UINT#1;
END_IF;
IF xStartCheckSafety THEN
	uiStartConditionsMet := uiStartConditionsMet + UINT#1;
END_IF;

xFaultAllowed := (eState = E_CELL_MANAGER_STATE.IDLE)
	AND NOT xRunning
	AND NOT xGlobalError
	AND NOT xMotionBusy
	AND NOT stRobotStatus.xBusy
	AND NOT stMagazineStatus.xBusy
	AND NOT xAnyMachineBusy
	AND (Error.dwErrorActive = DWORD#0);
fbFaultInjector(Request := FaultRequest, xOwnerAllowed := xFaultAllowed);
FaultStatus := fbFaultInjector.Status;

IF fbFaultInjector.Status.xRejected THEN
	Diag.stWarning.uiCode := WRN_SIM_ERROR_NOT_ALLOWED;
	Diag.stWarning.udiSequence := Diag.stWarning.udiSequence + UDINT#1;
	IF Diag.stWarning.udiSequence = UDINT#0 THEN
		Diag.stWarning.udiSequence := UDINT#1;
	END_IF;
END_IF;

IF rtStart.Q
AND xSafetyHomeRequired
AND NOT xRobotAtSafetyHome
AND NOT (xRunning AND xStopRequested) THEN
	Diag.stWarning.uiCode := WRN_SAFETY_HOME_REQUIRED;
	Diag.stWarning.udiSequence := Diag.stWarning.udiSequence + UDINT#1;
	IF Diag.stWarning.udiSequence = UDINT#0 THEN
		Diag.stWarning.udiSequence := UDINT#1;
	END_IF;
ELSIF rtStart.Q AND NOT (xReadyToStart OR (xRunning AND xStopRequested)) THEN
	Diag.stWarning.uiCode := WRN_START_NOT_READY;
	Diag.stWarning.udiSequence := Diag.stWarning.udiSequence + UDINT#1;
	IF Diag.stWarning.udiSequence = UDINT#0 THEN
		Diag.stWarning.udiSequence := UDINT#1;
	END_IF;
END_IF;

IF rtStop.Q AND NOT xRunning THEN
	Diag.stWarning.uiCode := WRN_STOP_NOT_RUNNING;
	Diag.stWarning.udiSequence := Diag.stWarning.udiSequence + UDINT#1;
	IF Diag.stWarning.udiSequence = UDINT#0 THEN
		Diag.stWarning.udiSequence := UDINT#1;
	END_IF;
END_IF;

IF (uiModeRejectReason = UINT#2) OR (uiModeRejectReason = UINT#3) THEN
	IF uiModeRejectReason = UINT#2 THEN
		Diag.stWarning.uiCode := WRN_MANUAL_MODE_REJECTED;
	ELSE
		Diag.stWarning.uiCode := WRN_AUTOMATIC_MODE_REJECTED;
	END_IF;
	Diag.stWarning.udiSequence := Diag.stWarning.udiSequence + UDINT#1;
	IF Diag.stWarning.udiSequence = UDINT#0 THEN
		Diag.stWarning.udiSequence := UDINT#1;
	END_IF;
END_IF;

// Ответы HMI принимаются только пока PLC явно публикует активный шаг опроса.
xOperatorPromptState := (eState = E_CELL_MANAGER_STATE.WAIT_GRIPPER1_CONTENT)
	OR (eState = E_CELL_MANAGER_STATE.WAIT_GRIPPER1_TYPE)
	OR (eState = E_CELL_MANAGER_STATE.WAIT_GRIPPER2_CONTENT)
	OR (eState = E_CELL_MANAGER_STATE.WAIT_GRIPPER2_TYPE)
	OR (eState = E_CELL_MANAGER_STATE.WAIT_START_MACHINE);
xOperatorChoiceAllowed := xOperatorPromptState
	AND NOT xManual
	AND NOT xGlobalError
	AND (Error.dwErrorActive = DWORD#0)
	AND xRobotInterfaceReady
	AND xConfigurationValid
	AND xPointsConfigured
	AND xDrivesReady
	AND xRobotReady
	AND xMagazineReady
	AND (NOT xSafetyHomeRequired OR xRobotAtSafetyHome);
// Отмена не должна блокироваться из-за временно потерянной готовности:
// оператор всегда может закрыть незавершённый предпусковой опрос.
xOperatorCancelAllowed := xOperatorPromptState;

IF rtOperatorChoice.Q AND NOT xOperatorChoiceAllowed THEN
	Diag.stWarning.uiCode := WRN_OPERATOR_REPLY_REJECTED;
	Diag.stWarning.udiSequence := Diag.stWarning.udiSequence + UDINT#1;
	IF Diag.stWarning.udiSequence = UDINT#0 THEN
		Diag.stWarning.udiSequence := UDINT#1;
	END_IF;
END_IF;

IF rtOperatorCancel.Q THEN
	IF xOperatorCancelAllowed THEN
		uiBlankPayloadType := UINT#0;
		uiDetailPayloadType := UINT#0;
		uiSelectedMachine := UINT#0;
		uiSelectedType := UINT#0;
		eMachineOperation := E_MACHINE_OPERATION.NONE;
		eState := E_CELL_MANAGER_STATE.IDLE;
	ELSE
		Diag.stWarning.uiCode := WRN_OPERATOR_CANCEL_REJECTED;
		Diag.stWarning.udiSequence := Diag.stWarning.udiSequence + UDINT#1;
		IF Diag.stWarning.udiSequence = UDINT#0 THEN
			Diag.stWarning.udiSequence := UDINT#1;
		END_IF;
	END_IF;
END_IF;

// Если оператор или внешний контроллер изменил захваты во время вопроса, старый ответ больше недостоверен.
IF xOperatorPromptState
AND NOT rtOperatorCancel.Q
AND ((stRobotStatus.xBlankAvailable <> xPrestartGripper1Occupied)
	OR (stRobotStatus.xDetailAvailable <> xPrestartGripper2Occupied)) THEN
	Diag.stWarning.uiCode := WRN_OPERATOR_REPLY_REJECTED;
	Diag.stWarning.udiSequence := Diag.stWarning.udiSequence + UDINT#1;
	IF Diag.stWarning.udiSequence = UDINT#0 THEN
		Diag.stWarning.udiSequence := UDINT#1;
	END_IF;
	uiBlankPayloadType := UINT#0;
	uiDetailPayloadType := UINT#0;
	eState := E_CELL_MANAGER_STATE.IDLE;
END_IF;

IF xOperatorPromptState
AND xManual THEN
	uiBlankPayloadType := UINT#0;
	uiDetailPayloadType := UINT#0;
	uiSelectedMachine := UINT#0;
	uiSelectedType := UINT#0;
	eMachineOperation := E_MACHINE_OPERATION.NONE;
	eState := E_CELL_MANAGER_STATE.IDLE;
END_IF;

// Условия ожидания не являются ошибкой и не останавливают ячейку. Каждое
// предупреждение регистрируется один раз на непрерывный эпизод; после очистки
// причины новое появление условия создаст новую запись журнала.
IF xNoDetailDestinationCondition
AND NOT xDetailDestinationWarningActive THEN
	Diag.stWarning.uiCode := WRN_NO_DETAIL_DESTINATION;
	Diag.stWarning.udiSequence := Diag.stWarning.udiSequence + UDINT#1;
	IF Diag.stWarning.udiSequence = UDINT#0 THEN
		Diag.stWarning.udiSequence := UDINT#1;
	END_IF;
END_IF;
xDetailDestinationWarningActive := xNoDetailDestinationCondition;

IF xNoBlankStockCondition
AND NOT xBlankStockWarningActive THEN
	Diag.stWarning.uiCode := WRN_NO_BLANK_STOCK;
	Diag.stWarning.udiSequence := Diag.stWarning.udiSequence + UDINT#1;
	IF Diag.stWarning.udiSequence = UDINT#0 THEN
		Diag.stWarning.udiSequence := UDINT#1;
	END_IF;
END_IF;
xBlankStockWarningActive := xNoBlankStockCondition;

IF rtStop.Q OR xManual THEN
	xStopRequested := TRUE;
ELSIF rtStart.Q AND xRunning
AND (eState <> E_CELL_MANAGER_STATE.MACHINE_FAULT_STOP) THEN
	xStopRequested := FALSE;
END_IF;

// Ошибка робота становится ошибкой автоматического цикла только когда ячейка
// действительно выполняет цикл. В IDLE ручная ошибка остаётся у своего
// первичного владельца (ось, группа или робот) и не создаёт ложный каскад.
IF xRunning AND stRobotStatus.xError THEN
	xSafetyHomeRequired := TRUE;
	xStoppedPoseValid := FALSE;
	Error.dwErrorActive := Error.dwErrorActive OR ERR_ROBOT;
	eState := E_CELL_MANAGER_STATE.ERROR;
END_IF;

IF xGlobalError
AND (eState <> E_CELL_MANAGER_STATE.IDLE)
AND (eState <> E_CELL_MANAGER_STATE.ERROR) THEN
	// Не каждая общая авария требует возврата. Защёлкиваем только ситуацию,
	// где прервано движение либо робот мог находиться внутри станка/магазина.
	IF stRobotStatus.xBusy
	OR xMotionBusy
	OR (eState = E_CELL_MANAGER_STATE.ROUTE_TO_TARGET)
	OR (eState = E_CELL_MANAGER_STATE.RELEASE_ROBOT_COMMAND)
	OR (eState = E_CELL_MANAGER_STATE.SERVICE_TARGET)
	OR (eState = E_CELL_MANAGER_STATE.MAGAZINE_EXECUTE)
	OR (eState = E_CELL_MANAGER_STATE.RELEASE_MAGAZINE)
	OR (eState = E_CELL_MANAGER_STATE.MACHINE_FAULT_STOP) THEN
		xSafetyHomeRequired := TRUE;
		xStoppedPoseValid := FALSE;
	END_IF;
	Error.dwErrorActive := Error.dwErrorActive OR ERR_GLOBAL_STOP;
	eState := E_CELL_MANAGER_STATE.ERROR;
END_IF;

// Штатный Stop ждёт безопасную технологическую границу. Тестовый Abort ждать
// её не должен: удерживаем Stop владельцев и не даём автоматам выдать новую
// команду, пока Motion фактически не закончил торможение.
IF xTestAbort THEN
	eState := E_CELL_MANAGER_STATE.TEST_ABORT_STOP;
END_IF;

// При передаче I/O оператору нельзя ждать программные Busy: именно зависший
// владелец может требовать восстановления. Аварии и физический груз сохраняются.
IF xIoManual THEN
	xRunning := FALSE;
	xStopRequested := FALSE;
	xMachineServiceStarted := FALSE;
	xReselectAfterRobotRelease := FALSE;
	xSafetyHomeRequired := TRUE;
	xStoppedPoseValid := FALSE;
	uiSelectedMachine := UINT#0;
	uiSelectedType := UINT#0;
	eMachineOperation := E_MACHINE_OPERATION.NONE;
	eMagazineOperation := E_MAGAZINE_OPERATION.NONE;
	iTakeSlot := SINT#0;
	iPutSlot := SINT#0;
	iTakeOriginSlot := SINT#0;
	FOR uiMachine := FIRST_MACHINE TO LAST_MACHINE DO
		axMachineStartPending[uiMachine] := FALSE;
	END_FOR;
	// Передача I/O оператору отменяет внутреннюю привязку прежнего цикла.
	uiReturnMagazine := UINT#0;
	uiSupplyMagazine := UINT#0;
	IF eState <> E_CELL_MANAGER_STATE.ERROR THEN
		eState := E_CELL_MANAGER_STATE.IDLE;
	END_IF;
END_IF;

// ГК не зависит от готовности палет. Если магазин потерян после выгрузки,
// сначала доставляем вызванную деталь на свободный ГК либо паркуемся у занятого.
IF xRunning AND xGeometryHeld AND stRobotStatus.xDetailAvailable
AND (eState = E_CELL_MANAGER_STATE.WAIT_MAGAZINE)
AND NOT stRobotStatus.xBusy AND NOT xMotionBusy THEN
	PlanGeometry();
END_IF;

CASE eState OF
	E_CELL_MANAGER_STATE.IDLE:
		xRunning := FALSE;
		xStopRequested := FALSE;
		xMachineServiceStarted := FALSE;
		xReselectAfterRobotRelease := FALSE;
		eMagazineOperation := E_MAGAZINE_OPERATION.NONE;
		IF fbFaultInjector.xBothGrippers THEN
			Error.dwErrorActive := Error.dwErrorActive OR ERR_BOTH_GRIPPERS;
			eState := E_CELL_MANAGER_STATE.ERROR;
		ELSIF rtStart.Q AND NOT xManual THEN
			IF xReadyToStart THEN
				xPrestartGripper1Occupied := stRobotStatus.xBlankAvailable;
				xPrestartGripper2Occupied := stRobotStatus.xDetailAvailable;
				uiBlankPayloadType := UINT#0;
				uiDetailPayloadType := UINT#0;
				uiSelectedMachine := UINT#0;
				uiSelectedType := UINT#0;
				eMachineOperation := E_MACHINE_OPERATION.NONE;
				// Новый Start заново идентифицирует уже находящийся в захвате груз.
				// Слот происхождения прошлого цикла к нему не относится: иначе
				// RETURN_BLANK может попытаться положить груз в занятый чужой слот.
				iTakeSlot := SINT#0;
				iPutSlot := SINT#0;
				iTakeOriginSlot := SINT#0;
				eState := E_CELL_MANAGER_STATE.PRESTART_IDENTIFY;
				uiReturnMagazine := UINT#0;
				uiSupplyMagazine := UINT#0;
			END_IF;
		END_IF;

	E_CELL_MANAGER_STATE.PRESTART_IDENTIFY:
		IF xManual THEN
			eState := E_CELL_MANAGER_STATE.IDLE;
		ELSIF xPrestartGripper1Occupied THEN
			eState := E_CELL_MANAGER_STATE.WAIT_GRIPPER1_CONTENT;
		ELSIF xPrestartGripper2Occupied THEN
			eState := E_CELL_MANAGER_STATE.WAIT_GRIPPER2_CONTENT;
		ELSE
			xSafetyHomeRequired := FALSE;
			xStoppedPoseValid := FALSE;
			xRunning := TRUE;
			eState := E_CELL_MANAGER_STATE.PLAN_TARGET;
		END_IF;

	E_CELL_MANAGER_STATE.WAIT_GRIPPER1_CONTENT:
		IF rtOperatorChoice.Q AND xOperatorChoiceAllowed THEN
			IF uiOperatorChoice = UINT#1 THEN
				IF Config.uiTypeCount = UINT#1 THEN
					uiBlankPayloadType := UINT#1;
					IF xPrestartGripper2Occupied THEN
						eState := E_CELL_MANAGER_STATE.WAIT_GRIPPER2_CONTENT;
					ELSE
						xSafetyHomeRequired := FALSE;
						xStoppedPoseValid := FALSE;
						xRunning := TRUE;
						eState := E_CELL_MANAGER_STATE.PLAN_TARGET;
					END_IF;
				ELSE
					eState := E_CELL_MANAGER_STATE.WAIT_GRIPPER1_TYPE;
				END_IF;
			ELSIF uiOperatorChoice = UINT#2 THEN
				Diag.stWarning.uiCode := WRN_GRIPPER1_CONTENT;
				Diag.stWarning.udiSequence := Diag.stWarning.udiSequence + UDINT#1;
				IF Diag.stWarning.udiSequence = UDINT#0 THEN Diag.stWarning.udiSequence := UDINT#1; END_IF;
				eState := E_CELL_MANAGER_STATE.IDLE;
			ELSE
				Diag.stWarning.uiCode := WRN_OPERATOR_REPLY_REJECTED;
				Diag.stWarning.udiSequence := Diag.stWarning.udiSequence + UDINT#1;
				IF Diag.stWarning.udiSequence = UDINT#0 THEN Diag.stWarning.udiSequence := UDINT#1; END_IF;
				eState := E_CELL_MANAGER_STATE.IDLE;
			END_IF;
		END_IF;

	E_CELL_MANAGER_STATE.WAIT_GRIPPER1_TYPE:
		IF rtOperatorChoice.Q AND xOperatorChoiceAllowed THEN
			IF (uiOperatorChoice >= UINT#1)
			AND (uiOperatorChoice <= Config.uiTypeCount) THEN
				uiBlankPayloadType := uiOperatorChoice;
				IF xPrestartGripper2Occupied THEN
					eState := E_CELL_MANAGER_STATE.WAIT_GRIPPER2_CONTENT;
				ELSE
					xSafetyHomeRequired := FALSE;
					xStoppedPoseValid := FALSE;
					xRunning := TRUE;
					eState := E_CELL_MANAGER_STATE.PLAN_TARGET;
				END_IF;
			ELSE
				Diag.stWarning.uiCode := WRN_PAYLOAD_TYPE_CHOICE;
				Diag.stWarning.udiSequence := Diag.stWarning.udiSequence + UDINT#1;
				IF Diag.stWarning.udiSequence = UDINT#0 THEN Diag.stWarning.udiSequence := UDINT#1; END_IF;
				eState := E_CELL_MANAGER_STATE.IDLE;
			END_IF;
		END_IF;

	E_CELL_MANAGER_STATE.WAIT_GRIPPER2_CONTENT:
		IF rtOperatorChoice.Q AND xOperatorChoiceAllowed THEN
			IF uiOperatorChoice = UINT#2 THEN
				IF Config.uiTypeCount = UINT#1 THEN
					uiDetailPayloadType := UINT#1;
				ELSE
					eState := E_CELL_MANAGER_STATE.WAIT_GRIPPER2_TYPE;
				END_IF;
				IF (Config.uiTypeCount = UINT#1) AND xPrestartGripper1Occupied THEN
					IF uiOperatorMachineMask <> UINT#0 THEN
						eState := E_CELL_MANAGER_STATE.WAIT_START_MACHINE;
					ELSE
						// Нет пустого совместимого станка: это не тупик. После
						// идентификации обоих грузов планировщик сначала уложит деталь.
						xSafetyHomeRequired := FALSE;
						xStoppedPoseValid := FALSE;
						xRunning := TRUE;
						eState := E_CELL_MANAGER_STATE.PLAN_TARGET;
					END_IF;
				ELSIF Config.uiTypeCount = UINT#1 THEN
					xSafetyHomeRequired := FALSE;
					xStoppedPoseValid := FALSE;
					xRunning := TRUE;
					eState := E_CELL_MANAGER_STATE.PLAN_TARGET;
				END_IF;
			ELSIF uiOperatorChoice = UINT#1 THEN
				Diag.stWarning.uiCode := WRN_GRIPPER2_CONTENT;
				Diag.stWarning.udiSequence := Diag.stWarning.udiSequence + UDINT#1;
				IF Diag.stWarning.udiSequence = UDINT#0 THEN Diag.stWarning.udiSequence := UDINT#1; END_IF;
				eState := E_CELL_MANAGER_STATE.IDLE;
			ELSE
				Diag.stWarning.uiCode := WRN_OPERATOR_REPLY_REJECTED;
				Diag.stWarning.udiSequence := Diag.stWarning.udiSequence + UDINT#1;
				IF Diag.stWarning.udiSequence = UDINT#0 THEN Diag.stWarning.udiSequence := UDINT#1; END_IF;
				eState := E_CELL_MANAGER_STATE.IDLE;
			END_IF;
		END_IF;

	E_CELL_MANAGER_STATE.WAIT_GRIPPER2_TYPE:
		IF rtOperatorChoice.Q AND xOperatorChoiceAllowed THEN
			IF (uiOperatorChoice >= UINT#1)
			AND (uiOperatorChoice <= Config.uiTypeCount) THEN
				uiDetailPayloadType := uiOperatorChoice;
				IF xPrestartGripper1Occupied THEN
					IF uiOperatorMachineMask <> UINT#0 THEN
						eState := E_CELL_MANAGER_STATE.WAIT_START_MACHINE;
					ELSE
						xSafetyHomeRequired := FALSE;
						xStoppedPoseValid := FALSE;
						xRunning := TRUE;
						eState := E_CELL_MANAGER_STATE.PLAN_TARGET;
					END_IF;
				ELSE
					xSafetyHomeRequired := FALSE;
					xStoppedPoseValid := FALSE;
					xRunning := TRUE;
					eState := E_CELL_MANAGER_STATE.PLAN_TARGET;
				END_IF;
			ELSE
				Diag.stWarning.uiCode := WRN_PAYLOAD_TYPE_CHOICE;
				Diag.stWarning.udiSequence := Diag.stWarning.udiSequence + UDINT#1;
				IF Diag.stWarning.udiSequence = UDINT#0 THEN Diag.stWarning.udiSequence := UDINT#1; END_IF;
				eState := E_CELL_MANAGER_STATE.IDLE;
			END_IF;
		END_IF;

	E_CELL_MANAGER_STATE.WAIT_START_MACHINE:
		IF (uiDetailPayloadType < UINT#1)
		OR (uiDetailPayloadType > Config.uiTypeCount) THEN
			Diag.stWarning.uiCode := WRN_PAYLOAD_TYPE_CHOICE;
			Diag.stWarning.udiSequence := Diag.stWarning.udiSequence + UDINT#1;
			IF Diag.stWarning.udiSequence = UDINT#0 THEN Diag.stWarning.udiSequence := UDINT#1; END_IF;
			eState := E_CELL_MANAGER_STATE.IDLE;
		ELSIF stMagazineStatus.stTypeStatus.aiFreeSlot[uiDetailPayloadType] = SINT#0 THEN
			Diag.stWarning.uiCode := WRN_DETAIL_SLOT_REQUIRED;
			Diag.stWarning.udiSequence := Diag.stWarning.udiSequence + UDINT#1;
			IF Diag.stWarning.udiSequence = UDINT#0 THEN Diag.stWarning.udiSequence := UDINT#1; END_IF;
			eState := E_CELL_MANAGER_STATE.IDLE;
		ELSIF uiOperatorMachineMask = UINT#0 THEN
			// Пока оператор отвечал, пустой станок мог стать недоступен. Сохраняем
			// оба груза и передаём решение общему планировщику вместо отмены старта.
			xSafetyHomeRequired := FALSE;
			xStoppedPoseValid := FALSE;
			xRunning := TRUE;
			eState := E_CELL_MANAGER_STATE.PLAN_TARGET;
		ELSIF rtOperatorChoice.Q AND xOperatorChoiceAllowed THEN
			IF ((uiOperatorChoice = UINT#1) AND ((uiOperatorMachineMask AND UINT#1) <> UINT#0))
			OR ((uiOperatorChoice = UINT#2) AND ((uiOperatorMachineMask AND UINT#2) <> UINT#0))
			OR ((uiOperatorChoice = UINT#3) AND ((uiOperatorMachineMask AND UINT#4) <> UINT#0)) THEN
				uiSelectedMachine := uiOperatorChoice;
				uiSelectedType := uiBlankPayloadType;
				eMachineOperation := E_MACHINE_OPERATION.LOAD;
				xSafetyHomeRequired := FALSE;
				xStoppedPoseValid := FALSE;
				xRunning := TRUE;
				eState := E_CELL_MANAGER_STATE.ROUTE_TO_TARGET;
			ELSE
				Diag.stWarning.uiCode := WRN_START_MACHINE_CHOICE;
				Diag.stWarning.udiSequence := Diag.stWarning.udiSequence + UDINT#1;
				IF Diag.stWarning.udiSequence = UDINT#0 THEN Diag.stWarning.udiSequence := UDINT#1; END_IF;
				eState := E_CELL_MANAGER_STATE.IDLE;
			END_IF;
		END_IF;

	E_CELL_MANAGER_STATE.PLAN_TARGET:
		IF xStopRequested
		AND NOT stRobotStatus.xBusy
		AND NOT stMagazineStatus.xBusy THEN
			xRunning := FALSE;
			eState := E_CELL_MANAGER_STATE.IDLE;

		ELSIF PlanGeometry() THEN
			// Метод зафиксировал резерв или безопасное ожидание свободного ГК.
		ELSIF stRobotStatus.xBlankAvailable
		AND stRobotStatus.xDetailAvailable THEN
			// Два груза после аварийного восстановления — штатная ситуация. Сначала
			// ищем пустой готовый станок строго по типу заготовки. Если загрузить её
			// прямо сейчас некуда, освобождаем захват 2 операцией PUT.
			IF (uiBlankPayloadType < UINT#1)
			OR (uiBlankPayloadType > Config.uiTypeCount) THEN
				Error.dwErrorActive := Error.dwErrorActive OR ERR_MAGAZINE;
				eState := E_CELL_MANAGER_STATE.ERROR;
			ELSIF (uiDetailPayloadType < UINT#1)
			OR (uiDetailPayloadType > Config.uiTypeCount) THEN
				Error.dwErrorActive := Error.dwErrorActive OR ERR_MACHINE;
				eState := E_CELL_MANAGER_STATE.ERROR;
			ELSE
				uiCandidateMachine := UINT#0;
				FOR uiMachine := FIRST_MACHINE TO LAST_MACHINE DO
					IF (uiCandidateMachine = UINT#0)
					AND IsMachineCompatible(
						uiMachine := uiMachine,
						uiProductType := uiBlankPayloadType
					)
					AND astMachineStatus[uiMachine].xCanAcceptService
					AND (astMachineStatus[uiMachine].ePartState = E_PART_STATE.EMPTY) THEN
						uiCandidateMachine := uiMachine;
					END_IF;
				END_FOR;

				IF uiCandidateMachine > UINT#0 THEN
					uiSelectedMachine := uiCandidateMachine;
					uiSelectedType := uiBlankPayloadType;
					eMachineOperation := E_MACHINE_OPERATION.LOAD;
					xMachineServiceStarted := FALSE;
					eState := E_CELL_MANAGER_STATE.ROUTE_TO_TARGET;
				ELSIF (stMagazineStatus.stTypeStatus.aiFreeSlot[uiDetailPayloadType] > SINT#0)
				AND xMagazineReady THEN
					uiSelectedMachine := UINT#0;
					uiSelectedType := UINT#0;
					eMachineOperation := E_MACHINE_OPERATION.NONE;
					iTakeSlot := SINT#0;
					iTakeOriginSlot := SINT#0;
					iPutSlot := stMagazineStatus.stTypeStatus.aiFreeSlot[uiDetailPayloadType];
					eMagazineOperation := E_MAGAZINE_OPERATION.PUT;
					eState := E_CELL_MANAGER_STATE.MAGAZINE_EXECUTE;
				ELSE
					eState := E_CELL_MANAGER_STATE.WAIT_MAGAZINE;
				END_IF;
			END_IF;

		ELSIF stRobotStatus.xBlankAvailable THEN
			IF (uiBlankPayloadType < UINT#1)
			OR (uiBlankPayloadType > Config.uiTypeCount) THEN
				Error.dwErrorActive := Error.dwErrorActive OR ERR_MAGAZINE;
				eState := E_CELL_MANAGER_STATE.ERROR;
			ELSE
				uiSelectedType := uiBlankPayloadType;
				uiCandidateMachine := SelectMachineForHeldBlank(
					uiProductType := uiBlankPayloadType,
					uiCurrentMachine := uiSelectedMachine
				);
				IF uiCandidateMachine > UINT#0 THEN
					uiSelectedMachine := uiCandidateMachine;
					eState := E_CELL_MANAGER_STATE.ROUTE_TO_TARGET;
				ELSE
					uiSelectedMachine := UINT#0;
					eState := E_CELL_MANAGER_STATE.SELECT_FALLBACK;
				END_IF;
			END_IF;

		ELSIF stRobotStatus.xDetailAvailable THEN
			uiBlankPayloadType := UINT#0;
			IF (uiDetailPayloadType < UINT#1)
			OR (uiDetailPayloadType > Config.uiTypeCount) THEN
				Error.dwErrorActive := Error.dwErrorActive OR ERR_MACHINE;
				eState := E_CELL_MANAGER_STATE.ERROR;
			ELSIF NOT xMagazineReady THEN
				eState := E_CELL_MANAGER_STATE.WAIT_MAGAZINE;
			ELSE
				// При полной палете CHANGE сначала освобождает слот взятием заготовки.
				// Станок назначения может быть пустым, готовым к обмену или обрабатывать.
				iPutSlot := stMagazineStatus.stTypeStatus.aiFreeSlot[uiDetailPayloadType];
				uiCandidateMachine := SelectMachineBeforeTake();
				uiSelectedMachine := UINT#0;
				uiSelectedType := UINT#0;
				iTakeSlot := SINT#0;
				iTakeOriginSlot := SINT#0;
				eMachineOperation := E_MACHINE_OPERATION.NONE;

				// Закрытый или переходный первый захват исключает CHANGE, даже если
				// логический флаг груза сейчас снят.
				IF stRobotStatus.xGripper1Open
				AND ((uiReturnMagazine = UINT#0) OR (uiReturnMagazine = uiActiveMagazine))
				AND (uiCandidateMachine >= FIRST_MACHINE)
				AND (uiCandidateMachine <= LAST_MACHINE) THEN
					uiSelectedMachine := uiCandidateMachine;
					uiSelectedType := Config.auiMachineType[uiSelectedMachine];
					IF (uiSelectedType >= UINT#1)
					AND (uiSelectedType <= Config.uiTypeCount) THEN
						iTakeSlot := stMagazineStatus.stTypeStatus.aiBlankSlot[uiSelectedType];
					END_IF;
				END_IF;

				// Индексы проверяются до обращения к карте секций. Обычный AND в
				// CODESYS не используется как защита динамического индекса массива.
				IF iPutSlot = SINT#0 THEN
					iPutSlot := iTakeSlot;
				END_IF;
				IF (iPutSlot >= SINT#1)
				AND (SINT_TO_UINT(iPutSlot) <= SINT_TO_UINT(GVL_CELL_SETTINGS.NumberDetail))
				AND (iTakeSlot >= SINT#1)
				AND (SINT_TO_UINT(iTakeSlot) <= SINT_TO_UINT(GVL_CELL_SETTINGS.NumberDetail)) THEN
					xChangePrepared := TRUE;
				END_IF;

				IF xChangePrepared THEN
					iTakeOriginSlot := iTakeSlot;
					eMagazineOperation := E_MAGAZINE_OPERATION.CHANGE;
					eState := E_CELL_MANAGER_STATE.MAGAZINE_EXECUTE;
				ELSE
					// Если следующую заготовку нельзя безопасно назначить, сначала
					// освобождаем второй захват и пересчитываем маршрут после PUT.
					uiSelectedMachine := UINT#0;
					uiSelectedType := UINT#0;
					iTakeSlot := SINT#0;
					iTakeOriginSlot := SINT#0;
					IF stMagazineStatus.stTypeStatus.aiFreeSlot[uiDetailPayloadType] > SINT#0 THEN
						iPutSlot := stMagazineStatus.stTypeStatus.aiFreeSlot[uiDetailPayloadType];
						eMagazineOperation := E_MAGAZINE_OPERATION.PUT;
						eState := E_CELL_MANAGER_STATE.MAGAZINE_EXECUTE;
					ELSE
						iPutSlot := SINT#0;
						eMagazineOperation := E_MAGAZINE_OPERATION.NONE;
						eState := E_CELL_MANAGER_STATE.WAIT_MAGAZINE;
					END_IF;
				END_IF;
			END_IF;

		ELSE
			uiBlankPayloadType := UINT#0;
			uiDetailPayloadType := UINT#0;
			uiCandidateMachine := SelectMachineBeforeTake();
			IF uiCandidateMachine > UINT#0 THEN
				IF NOT xMagazineReady THEN
					eState := E_CELL_MANAGER_STATE.WAIT_MAGAZINE;
				ELSE
					uiSelectedMachine := uiCandidateMachine;
					uiSelectedType := Config.auiMachineType[uiSelectedMachine];
					iTakeSlot := stMagazineStatus.stTypeStatus.aiBlankSlot[uiSelectedType];
					iTakeOriginSlot := iTakeSlot;
					iPutSlot := SINT#0;
					eMachineOperation := E_MACHINE_OPERATION.NONE;
					eMagazineOperation := E_MAGAZINE_OPERATION.TAKE;
					eState := E_CELL_MANAGER_STATE.MAGAZINE_EXECUTE;
				END_IF;
			ELSE
				// Заготовок в магазине нет — выбираем готовую деталь для отдельной выгрузки.
				uiCandidateMachine := SelectMachineForUnload(uiCurrentMachine := UINT#0);
				IF uiCandidateMachine > UINT#0 THEN
					uiSelectedMachine := uiCandidateMachine;
					uiSelectedType := Config.auiMachineType[uiSelectedMachine];
					eMachineOperation := E_MACHINE_OPERATION.UNLOAD;
					xMachineServiceStarted := FALSE;
					iTakeSlot := SINT#0;
					iPutSlot := SINT#0;
					IF xMagazineReady THEN
						eState := E_CELL_MANAGER_STATE.ROUTE_TO_TARGET;
					ELSE
						eState := E_CELL_MANAGER_STATE.WAIT_MAGAZINE;
					END_IF;
				ELSE
					IF stMagazineStatus.xFinished THEN
						eState := E_CELL_MANAGER_STATE.WAIT_MAGAZINE;
					ELSE
						eState := E_CELL_MANAGER_STATE.WAIT_TARGET;
					END_IF;
				END_IF;
			END_IF;
		END_IF;

	E_CELL_MANAGER_STATE.MAGAZINE_EXECUTE:
		IF xGeometryHeld AND (uiGeometryMachine >= UINT#1) AND (uiGeometryMachine <= UINT#3)
		AND (stMagazineStatus.udiProducedPartsTotal <> udiGeometryMagazineCounter)
		AND NOT stRobotStatus.xDetailAvailable AND stRobotStatus.xGripper2Open THEN
			GVL_GEOMETRY_CONTROL.astCalls[uiGeometryMachine].uiState := UINT#5;
			GVL_GEOMETRY_CONTROL.astCalls[uiGeometryMachine].uiReason := uiGeometryBypassReason;
			GVL_GEOMETRY_CONTROL.astCalls[uiGeometryMachine].uiMagazine := uiActiveMagazine;
			GVL_GEOMETRY_CONTROL.astCalls[uiGeometryMachine].uiSlot := SINT_TO_UINT(iPutSlot);
			IF GVL_TWO_PALLET.uiMode = UINT#1 THEN
				GVL_GEOMETRY_CONTROL.astCalls[uiGeometryMachine].uiPallet := GVL_TWO_PALLET.astStatus[uiActiveMagazine].uiRobotPallet;
			END_IF;
			F_GEOMETRY_EVENT(Call := GVL_GEOMETRY_CONTROL.astCalls[uiGeometryMachine]);
			GVL_GEOMETRY_CONTROL.stCellWarning.uiCode := UINT#50;
			GVL_GEOMETRY_CONTROL.stCellWarning.udiSequence := GVL_GEOMETRY_CONTROL.stCellWarning.udiSequence + UDINT#1;
			xGeometryHeld := FALSE; uiGeometryMachine := UINT#0;
		END_IF;
		Command.stMagazine.xExecute := TRUE;
		IF (eMagazineOperation = E_MAGAZINE_OPERATION.NONE) THEN
			Error.dwErrorActive := Error.dwErrorActive OR ERR_MAGAZINE;
			eState := E_CELL_MANAGER_STATE.ERROR;
		END_IF;

		IF stMagazineStatus.xError THEN
			Command.stMagazine.xExecute := FALSE;
			IF stMagazineStatus.xRobotStopRequired THEN
				xSafetyHomeRequired := TRUE;
				xStoppedPoseValid := FALSE;
				Error.dwErrorActive := Error.dwErrorActive OR ERR_MAGAZINE;
				eState := E_CELL_MANAGER_STATE.ERROR;
			ELSE
				xRunning := FALSE;
				eState := E_CELL_MANAGER_STATE.IDLE;
			END_IF;
		ELSIF stRobotStatus.xError THEN
			Error.dwErrorActive := Error.dwErrorActive OR ERR_ROBOT;
			eState := E_CELL_MANAGER_STATE.ERROR;
		ELSIF stMagazineStatus.xDone THEN
			eState := E_CELL_MANAGER_STATE.RELEASE_MAGAZINE;
		END_IF;

	E_CELL_MANAGER_STATE.RELEASE_MAGAZINE:
		IF stMagazineStatus.xError THEN
			IF stMagazineStatus.xRobotStopRequired THEN
				xSafetyHomeRequired := TRUE;
				xStoppedPoseValid := FALSE;
				Error.dwErrorActive := Error.dwErrorActive OR ERR_MAGAZINE;
				eState := E_CELL_MANAGER_STATE.ERROR;
			ELSE
				xRunning := FALSE;
				eState := E_CELL_MANAGER_STATE.IDLE;
			END_IF;
		ELSIF NOT stMagazineStatus.xBusy
		AND NOT stMagazineStatus.xDone THEN
			CASE eMagazineOperation OF
				E_MAGAZINE_OPERATION.TAKE:
					uiBlankPayloadType := uiSelectedType;
					uiReturnMagazine := uiActiveMagazine;
					uiSupplyMagazine := uiActiveMagazine;
				E_MAGAZINE_OPERATION.PUT:
					uiDetailPayloadType := UINT#0;
					uiReturnMagazine := UINT#0;
				E_MAGAZINE_OPERATION.CHANGE:
					uiDetailPayloadType := UINT#0;
					uiBlankPayloadType := uiSelectedType;
					uiReturnMagazine := uiActiveMagazine;
					uiSupplyMagazine := uiActiveMagazine;
				E_MAGAZINE_OPERATION.RETURN_BLANK:
					uiBlankPayloadType := UINT#0;
					uiReturnMagazine := UINT#0;
					uiSelectedType := UINT#0;
					iTakeOriginSlot := SINT#0;
					iTakeSlot := SINT#0;
					iPutSlot := SINT#0;
			END_CASE;
			eMagazineOperation := E_MAGAZINE_OPERATION.NONE;
			eState := E_CELL_MANAGER_STATE.PLAN_TARGET;
		END_IF;

	E_CELL_MANAGER_STATE.ROUTE_TO_TARGET:
		IF eMachineOperation = E_MACHINE_OPERATION.UNLOAD THEN
			IF stRobotStatus.eCurrentPoint = astMachineStatus[uiSelectedMachine].eAbovePoint THEN
				eState := E_CELL_MANAGER_STATE.WAIT_TARGET;
			ELSE
				Command.stRobot.xExecute := TRUE;
				Command.stRobot.eAction := E_ROBOT_ACTION.MOVE_TO_POINT;
				Command.stRobot.eSetPoint := astMachineStatus[uiSelectedMachine].eAbovePoint;
				IF stRobotStatus.xDone THEN
					xReselectAfterRobotRelease := FALSE;
					eState := E_CELL_MANAGER_STATE.RELEASE_ROBOT_COMMAND;
				END_IF;
			END_IF;
		ELSE
			IF (uiSelectedMachine >= FIRST_MACHINE)
			AND (uiSelectedMachine <= LAST_MACHINE) THEN
				RaisePayloadRouteWarning(
					uiPayloadType := uiBlankPayloadType,
					uiDestinationType := Config.auiMachineType[uiSelectedMachine]
				);
			END_IF;
			IF NOT IsMachineCompatible(
				uiMachine := uiSelectedMachine,
				uiProductType := uiBlankPayloadType
			) THEN
				xReselectAfterRobotRelease := TRUE;
				eState := E_CELL_MANAGER_STATE.RELEASE_ROBOT_COMMAND;
			ELSIF stRobotStatus.eCurrentPoint = astMachineStatus[uiSelectedMachine].eAbovePoint THEN
				eState := E_CELL_MANAGER_STATE.WAIT_TARGET;
			ELSE
				Command.stRobot.xExecute := TRUE;
				Command.stRobot.eAction := E_ROBOT_ACTION.MOVE_TO_POINT;
				Command.stRobot.eSetPoint := astMachineStatus[uiSelectedMachine].eAbovePoint;
				IF stRobotStatus.xDone THEN
					xReselectAfterRobotRelease := FALSE;
					eState := E_CELL_MANAGER_STATE.RELEASE_ROBOT_COMMAND;
				END_IF;
			END_IF;
		END_IF;

	E_CELL_MANAGER_STATE.RELEASE_ROBOT_COMMAND:
		IF stRobotStatus.xError THEN
			Error.dwErrorActive := Error.dwErrorActive OR ERR_ROBOT;
			eState := E_CELL_MANAGER_STATE.ERROR;
		ELSIF NOT stRobotStatus.xBusy
		AND NOT stRobotStatus.xDone
		AND NOT xMotionBusy THEN
			IF eMachineOperation = E_MACHINE_OPERATION.UNLOAD THEN
				eState := E_CELL_MANAGER_STATE.WAIT_TARGET;
			ELSIF xReselectAfterRobotRelease THEN
				xReselectAfterRobotRelease := FALSE;
				eState := E_CELL_MANAGER_STATE.SELECT_FALLBACK;
			ELSIF IsMachineCompatible(
				uiMachine := uiSelectedMachine,
				uiProductType := uiBlankPayloadType
			) THEN
				eState := E_CELL_MANAGER_STATE.WAIT_TARGET;
			ELSE
				eState := E_CELL_MANAGER_STATE.SELECT_FALLBACK;
			END_IF;
		END_IF;

	E_CELL_MANAGER_STATE.WAIT_TARGET:
		IF xStopRequested
		AND NOT stRobotStatus.xBusy THEN
			xRunning := FALSE;
			eState := E_CELL_MANAGER_STATE.IDLE;
		ELSIF (eMachineOperation = E_MACHINE_OPERATION.UNLOAD)
		AND NOT stRobotStatus.xBlankAvailable
		AND NOT stRobotStatus.xDetailAvailable THEN
			uiCandidateMachine := SelectMachineForUnload(uiCurrentMachine := uiSelectedMachine);
			IF uiCandidateMachine = UINT#0 THEN
				uiSelectedMachine := UINT#0;
				uiSelectedType := UINT#0;
				eMachineOperation := E_MACHINE_OPERATION.NONE;
				IF stMagazineStatus.xFinished THEN
					eState := E_CELL_MANAGER_STATE.WAIT_MAGAZINE;
				ELSE
					eState := E_CELL_MANAGER_STATE.PLAN_TARGET;
				END_IF;
			ELSIF uiCandidateMachine <> uiSelectedMachine THEN
				uiSelectedMachine := uiCandidateMachine;
				uiSelectedType := Config.auiMachineType[uiSelectedMachine];
				eState := E_CELL_MANAGER_STATE.ROUTE_TO_TARGET;
			ELSIF stRobotStatus.eCurrentPoint <> astMachineStatus[uiSelectedMachine].eAbovePoint THEN
				eState := E_CELL_MANAGER_STATE.ROUTE_TO_TARGET;
			ELSIF astMachineStatus[uiSelectedMachine].xCanAcceptService
			AND astMachineStatus[uiSelectedMachine].xServiceRequired
			AND (astMachineStatus[uiSelectedMachine].ePartState = E_PART_STATE.LOADED)
			AND (astMachineStatus[uiSelectedMachine].ePartType = E_PART_TYPE.DETAIL) THEN
				xMachineServiceStarted := FALSE;
				eState := E_CELL_MANAGER_STATE.SERVICE_TARGET;
			END_IF;
		ELSIF stRobotStatus.xBlankAvailable
		AND stRobotStatus.xDetailAvailable THEN
			// Выбранная пустая цель могла стать недоступной по дороге. Обслуживаем
			// только всё ещё пустой совместимый станок; иначе перепланируем через PUT.
			IF (uiSelectedMachine >= FIRST_MACHINE)
			AND (uiSelectedMachine <= LAST_MACHINE) THEN
				IF IsMachineCompatible(
					uiMachine := uiSelectedMachine,
					uiProductType := uiBlankPayloadType
				)
				AND (stRobotStatus.eCurrentPoint = astMachineStatus[uiSelectedMachine].eAbovePoint)
				AND astMachineStatus[uiSelectedMachine].xCanAcceptService
				AND (astMachineStatus[uiSelectedMachine].ePartState = E_PART_STATE.EMPTY) THEN
					eMachineOperation := E_MACHINE_OPERATION.LOAD;
					xMachineServiceStarted := FALSE;
					eState := E_CELL_MANAGER_STATE.SERVICE_TARGET;
				ELSE
					eState := E_CELL_MANAGER_STATE.PLAN_TARGET;
				END_IF;
			ELSE
				eState := E_CELL_MANAGER_STATE.PLAN_TARGET;
			END_IF;
		ELSIF stRobotStatus.xBlankAvailable THEN
			uiCandidateMachine := SelectMachineForHeldBlank(
				uiProductType := uiBlankPayloadType,
				uiCurrentMachine := uiSelectedMachine
			);
			IF uiCandidateMachine = UINT#0 THEN
				eState := E_CELL_MANAGER_STATE.SELECT_FALLBACK;
			ELSIF uiCandidateMachine <> uiSelectedMachine THEN
				uiSelectedMachine := uiCandidateMachine;
				eState := E_CELL_MANAGER_STATE.ROUTE_TO_TARGET;
			ELSIF stRobotStatus.eCurrentPoint <> astMachineStatus[uiSelectedMachine].eAbovePoint THEN
				eState := E_CELL_MANAGER_STATE.ROUTE_TO_TARGET;
			ELSIF astMachineStatus[uiSelectedMachine].xCanAcceptService
			AND astMachineStatus[uiSelectedMachine].xServiceRequired THEN
				eMachineOperation := astMachineStatus[uiSelectedMachine].eRecommendedOperation;
				axMachineStartPending[uiSelectedMachine] := FALSE;
				xMachineServiceStarted := FALSE;
				eState := E_CELL_MANAGER_STATE.SERVICE_TARGET;
			END_IF;
		ELSIF stRobotStatus.xDetailAvailable THEN
			// Готовая деталь в захвате обслуживается через общий план PUT.
			eState := E_CELL_MANAGER_STATE.PLAN_TARGET;
		ELSE
			uiCandidateMachine := SelectMachineBeforeTake();
			IF uiCandidateMachine > UINT#0 THEN
				eState := E_CELL_MANAGER_STATE.PLAN_TARGET;
			ELSE
				// В магазине нет заготовки: ожидаем готовую деталь станка,
				// которую можно выгрузить в свободный слот.
				uiCandidateMachine := SelectMachineForUnload(uiCurrentMachine := uiSelectedMachine);
				IF uiCandidateMachine > UINT#0 THEN
					uiSelectedMachine := uiCandidateMachine;
					uiSelectedType := Config.auiMachineType[uiSelectedMachine];
					eMachineOperation := E_MACHINE_OPERATION.UNLOAD;
					xMachineServiceStarted := FALSE;
					iTakeSlot := SINT#0;
					iPutSlot := SINT#0;
					IF xMagazineReady THEN
						eState := E_CELL_MANAGER_STATE.ROUTE_TO_TARGET;
					ELSE
						eState := E_CELL_MANAGER_STATE.WAIT_MAGAZINE;
					END_IF;
				ELSIF stMagazineStatus.xFinished THEN
					eState := E_CELL_MANAGER_STATE.WAIT_MAGAZINE;
				END_IF;
			END_IF;
		END_IF;

	E_CELL_MANAGER_STATE.SERVICE_TARGET:
		IF (uiSelectedMachine < FIRST_MACHINE)
		OR (uiSelectedMachine > LAST_MACHINE) THEN
			Error.dwErrorActive := Error.dwErrorActive OR ERR_MACHINE;
			eState := E_CELL_MANAGER_STATE.ERROR;
		ELSIF NOT xMachineServiceStarted AND NOT astMachineStatus[uiSelectedMachine].xBusy
		AND (eMachineOperation <> E_MACHINE_OPERATION.LOAD)
		AND axGeometryUnloadBlocked[uiSelectedMachine] THEN
			// До запуска рецепта повторно проверяем наличие доступного свободного ГК.
			// Деталь остаётся в патроне; ищем другую работу без команды станку.
			eState := E_CELL_MANAGER_STATE.SELECT_FALLBACK;
		ELSIF NOT xMachineServiceStarted
		AND (eMachineOperation <> E_MACHINE_OPERATION.UNLOAD)
		AND NOT IsMachineCompatible(
			uiMachine := uiSelectedMachine,
			uiProductType := uiBlankPayloadType
		) THEN
			RaisePayloadRouteWarning(
				uiPayloadType := uiBlankPayloadType,
				uiDestinationType := Config.auiMachineType[uiSelectedMachine]
			);
			eState := E_CELL_MANAGER_STATE.SELECT_FALLBACK;
		ELSE
			IF NOT xMachineServiceStarted AND NOT stRobotStatus.xDetailAvailable THEN xGeometryDetailCounted := FALSE; END_IF;
			IF stRobotStatus.xDetailAvailable AND NOT xGeometryDetailCounted
			AND ((eMachineOperation = E_MACHINE_OPERATION.CHANGE) OR (eMachineOperation = E_MACHINE_OPERATION.UNLOAD)) THEN
				xGeometryHeld := F_GEOMETRY_TAKE_DETAIL(uiMachine := uiSelectedMachine, uiProductType := Config.auiMachineType[uiSelectedMachine]);
				IF xGeometryHeld THEN uiGeometryMachine := uiSelectedMachine; uiGeometryBypassReason := UINT#0; END_IF;
				xGeometryDetailCounted := TRUE;
			END_IF;
			// Тип детали передаётся в FB_ROBOT сразу после фактического закрытия
			// второго захвата, а не после полного выхода робота из станка.
			IF stRobotStatus.xDetailAvailable
			AND ((eMachineOperation = E_MACHINE_OPERATION.CHANGE)
				OR (eMachineOperation = E_MACHINE_OPERATION.UNLOAD)) THEN
				uiDetailPayloadType := Config.auiMachineType[uiSelectedMachine];
			END_IF;
			IF eMachineOperation <> E_MACHINE_OPERATION.UNLOAD THEN
				RaisePayloadRouteWarning(
					uiPayloadType := uiBlankPayloadType,
					uiDestinationType := Config.auiMachineType[uiSelectedMachine]
				);
			END_IF;
			Command.axMachineExecute[uiSelectedMachine] := TRUE;
			IF astMachineStatus[uiSelectedMachine].xBusy THEN
				xMachineServiceStarted := TRUE;
			END_IF;

			IF astMachineStatus[uiSelectedMachine].xServiceRejected THEN
				Command.axMachineExecute[uiSelectedMachine] := FALSE;
				xMachineServiceStarted := FALSE;
				eMachineOperation := E_MACHINE_OPERATION.NONE;
				xReselectAfterRobotRelease := TRUE;
				eState := E_CELL_MANAGER_STATE.RELEASE_ROBOT_COMMAND;
			ELSIF astMachineStatus[uiSelectedMachine].xError THEN
				Command.axMachineExecute[uiSelectedMachine] := FALSE;
				xMachineServiceStarted := FALSE;
				// ROBOT_STOP уже публикует сам станок и обрабатывает FB_ROBOT.
				// Локальная ошибка без робота просто исключает станок из маршрута.
				eMachineOperation := E_MACHINE_OPERATION.NONE;
				xReselectAfterRobotRelease := TRUE;
				eState := E_CELL_MANAGER_STATE.RELEASE_ROBOT_COMMAND;
			ELSIF stRobotStatus.xError THEN
				Error.dwErrorActive := Error.dwErrorActive OR ERR_ROBOT;
				eState := E_CELL_MANAGER_STATE.ERROR;
			ELSIF astMachineStatus[uiSelectedMachine].xRobotReleased THEN
				// Вызов мог прийти после взятия детали, пока робот ещё менял заготовку.
				// Последняя проверка — после подтверждённого выхода, до сброса станка.
				// Только state 1: F_GEOMETRY_TAKE_DETAIL не считает выгрузку повторно
				// и привязывает вызов своей детали независимо от вызовов других станков.
				IF NOT xGeometryHeld AND stRobotStatus.xDetailAvailable
				AND ((eMachineOperation = E_MACHINE_OPERATION.CHANGE)
					OR (eMachineOperation = E_MACHINE_OPERATION.UNLOAD))
				AND (GVL_GEOMETRY_CONTROL.astCalls[uiSelectedMachine].uiState = UINT#1) THEN
					xGeometryHeld := F_GEOMETRY_TAKE_DETAIL(uiMachine := uiSelectedMachine, uiProductType := Config.auiMachineType[uiSelectedMachine]);
					IF xGeometryHeld THEN uiGeometryMachine := uiSelectedMachine; uiGeometryBypassReason := UINT#0; END_IF;
				END_IF;
				IF (eMachineOperation = E_MACHINE_OPERATION.LOAD)
				OR (eMachineOperation = E_MACHINE_OPERATION.CHANGE) THEN
					axMachineStartPending[uiSelectedMachine] := TRUE;
				END_IF;
				uiBlankPayloadType := UINT#0;
				IF (eMachineOperation = E_MACHINE_OPERATION.CHANGE)
				OR (eMachineOperation = E_MACHINE_OPERATION.UNLOAD) THEN
					uiDetailPayloadType := Config.auiMachineType[uiSelectedMachine];
				END_IF;
				uiSelectedMachine := UINT#0;
				uiSelectedType := UINT#0;
				xMachineServiceStarted := FALSE;
				eMachineOperation := E_MACHINE_OPERATION.NONE;
				eState := E_CELL_MANAGER_STATE.PLAN_TARGET;
			END_IF;
		END_IF;

	E_CELL_MANAGER_STATE.MACHINE_FAULT_STOP:
		// Удерживаем штатную остановку до полного освобождения Motion-слоя.
		// Первичная MachineAlarm/Timeout остаётся активной только в FB_MACHINE.
		Command.stRobot.xStop := stRobotStatus.xBusy OR xMotionBusy;
		IF NOT stRobotStatus.xBusy AND NOT xMotionBusy THEN
			xRunning := FALSE;
			xStopRequested := FALSE;
			xMachineServiceStarted := FALSE;
			xReselectAfterRobotRelease := FALSE;
			IF (uiSelectedMachine >= FIRST_MACHINE)
			AND (uiSelectedMachine <= LAST_MACHINE) THEN
				axMachineStartPending[uiSelectedMachine] := FALSE;
			END_IF;
			uiSelectedMachine := UINT#0;
			uiSelectedType := UINT#0;
			eMachineOperation := E_MACHINE_OPERATION.NONE;
			eState := E_CELL_MANAGER_STATE.IDLE;
		END_IF;

	E_CELL_MANAGER_STATE.SELECT_FALLBACK:
		IF xStopRequested
		AND NOT stRobotStatus.xBusy
		AND NOT stMagazineStatus.xBusy THEN
			xRunning := FALSE;
			eState := E_CELL_MANAGER_STATE.IDLE;
		ELSIF stRobotStatus.xDetailAvailable THEN
			// RETURN_BLANK запрещён при занятом захвате 2. Общий план сначала
			// попробует другой пустой станок, затем освободит готовую деталь через PUT.
			eState := E_CELL_MANAGER_STATE.PLAN_TARGET;
		ELSIF NOT stRobotStatus.xBlankAvailable THEN
			// Отказ UNLOAD до захвата оставляет робот пустым. Старый тип
			// заготовки не является грузом и не создаёт ошибку магазина.
			uiSelectedMachine := UINT#0;
			uiSelectedType := UINT#0;
			uiBlankPayloadType := UINT#0;
			eMachineOperation := E_MACHINE_OPERATION.NONE;
			eMagazineOperation := E_MAGAZINE_OPERATION.NONE;
			eState := E_CELL_MANAGER_STATE.PLAN_TARGET;
		ELSIF (uiBlankPayloadType < UINT#1)
		OR (uiBlankPayloadType > Config.uiTypeCount) THEN
			Error.dwErrorActive := Error.dwErrorActive OR ERR_MAGAZINE;
			eState := E_CELL_MANAGER_STATE.ERROR;
		ELSE
			uiCandidateMachine := SelectMachineForHeldBlank(
				uiProductType := uiBlankPayloadType,
				uiCurrentMachine := uiSelectedMachine
			);
		END_IF;
		IF (eState = E_CELL_MANAGER_STATE.SELECT_FALLBACK)
		AND (uiCandidateMachine > UINT#0) THEN
			uiSelectedMachine := uiCandidateMachine;
			uiSelectedType := uiBlankPayloadType;
			eState := E_CELL_MANAGER_STATE.ROUTE_TO_TARGET;
		ELSIF eState = E_CELL_MANAGER_STATE.SELECT_FALLBACK THEN
			uiSelectedMachine := UINT#0;
			eMachineOperation := E_MACHINE_OPERATION.NONE;
			eMagazineOperation := E_MAGAZINE_OPERATION.NONE;
			iPutSlot := SINT#0;
			IF NOT CanReturnHeldBlank() THEN
				// Один тип либо нет полезной работы другого типа: сохраняем
				// заготовку. WAIT_MAGAZINE заново проверяет маршруты без Start.
				eState := E_CELL_MANAGER_STATE.WAIT_MAGAZINE;
			ELSE
				// Исходный слот гарантированно освободился после подтверждённой TAKE.
				IF (iTakeOriginSlot >= SINT#1)
				AND (SINT_TO_UINT(iTakeOriginSlot) <= SINT_TO_UINT(GVL_CELL_SETTINGS.NumberDetail)) THEN
					iPutSlot := iTakeOriginSlot;
				END_IF;
				IF iPutSlot = SINT#0 THEN
					iPutSlot := stMagazineStatus.stTypeStatus.aiFreeSlot[uiBlankPayloadType];
				END_IF;
				IF (iPutSlot > SINT#0) AND xMagazineReady THEN
					eMagazineOperation := E_MAGAZINE_OPERATION.RETURN_BLANK;
					eState := E_CELL_MANAGER_STATE.MAGAZINE_EXECUTE;
				ELSE
					eState := E_CELL_MANAGER_STATE.WAIT_MAGAZINE;
				END_IF;
			END_IF;
		END_IF;

	E_CELL_MANAGER_STATE.WAIT_MAGAZINE:
		IF xStopRequested
		AND NOT stMagazineStatus.xBusy
		AND NOT stRobotStatus.xBusy THEN
			xRunning := FALSE;
			eState := E_CELL_MANAGER_STATE.IDLE;
		ELSIF stMagazineStatus.xError THEN
			IF stMagazineStatus.xRobotStopRequired THEN
				Error.dwErrorActive := Error.dwErrorActive OR ERR_MAGAZINE;
				eState := E_CELL_MANAGER_STATE.ERROR;
			ELSE
				xRunning := FALSE;
				eState := E_CELL_MANAGER_STATE.IDLE;
			END_IF;
		ELSIF stRobotStatus.xBlankAvailable
		AND stRobotStatus.xDetailAvailable THEN
			IF (uiBlankPayloadType < UINT#1)
			OR (uiBlankPayloadType > Config.uiTypeCount) THEN
				Error.dwErrorActive := Error.dwErrorActive OR ERR_MAGAZINE;
				eState := E_CELL_MANAGER_STATE.ERROR;
			ELSIF (uiDetailPayloadType < UINT#1)
			OR (uiDetailPayloadType > Config.uiTypeCount) THEN
				Error.dwErrorActive := Error.dwErrorActive OR ERR_MACHINE;
				eState := E_CELL_MANAGER_STATE.ERROR;
			ELSIF (uiOperatorMachineMask <> UINT#0)
			OR ((stMagazineStatus.stTypeStatus.aiFreeSlot[uiDetailPayloadType] > SINT#0)
				AND xMagazineReady) THEN
				eState := E_CELL_MANAGER_STATE.PLAN_TARGET;
			END_IF;
		ELSIF stRobotStatus.xBlankAvailable THEN
			IF (uiBlankPayloadType < UINT#1)
			OR (uiBlankPayloadType > Config.uiTypeCount) THEN
				Error.dwErrorActive := Error.dwErrorActive OR ERR_MAGAZINE;
				eState := E_CELL_MANAGER_STATE.ERROR;
			ELSE
				IF (SelectMachineForHeldBlank(
					uiProductType := uiBlankPayloadType,
					uiCurrentMachine := uiSelectedMachine
				) > UINT#0)
				OR CanReturnHeldBlank() THEN
					eState := E_CELL_MANAGER_STATE.SELECT_FALLBACK;
				END_IF;
			END_IF;
		ELSIF stRobotStatus.xDetailAvailable THEN
			IF (uiDetailPayloadType < UINT#1)
			OR (uiDetailPayloadType > Config.uiTypeCount) THEN
				Error.dwErrorActive := Error.dwErrorActive OR ERR_MACHINE;
				eState := E_CELL_MANAGER_STATE.ERROR;
			ELSE
				IF ((stMagazineStatus.stTypeStatus.aiFreeSlot[uiDetailPayloadType] > SINT#0)
					OR xActiveMagazineCanExchangeDetail)
				AND xMagazineReady THEN
					eState := E_CELL_MANAGER_STATE.PLAN_TARGET;
				END_IF;
			END_IF;
		ELSE
			uiCandidateMachine := SelectMachineBeforeTake();
			IF uiCandidateMachine = UINT#0 THEN
				uiCandidateMachine := SelectMachineForUnload(uiCurrentMachine := uiSelectedMachine);
			END_IF;
			IF uiCandidateMachine > UINT#0 THEN
				IF xMagazineReady THEN
					eState := E_CELL_MANAGER_STATE.PLAN_TARGET;
				ELSE
					eState := E_CELL_MANAGER_STATE.WAIT_MAGAZINE;
				END_IF;
			END_IF;
		END_IF;

	E_CELL_MANAGER_STATE.GEOMETRY_WAIT_FREE,
	E_CELL_MANAGER_STATE.GEOMETRY_DELIVER,
	E_CELL_MANAGER_STATE.GEOMETRY_RELEASE_COMMAND:
		RunGeometryRoute();

	E_CELL_MANAGER_STATE.ERROR:
		xRunning := FALSE;
		IF stRobotStatus.xBusy THEN
			Command.stRobot.xStop := TRUE;
		END_IF;
		IF stMagazineStatus.xBusy THEN
			Command.stMagazine.xStop := TRUE;
		END_IF;
		xResetAllowed := NOT xGlobalError
			AND NOT stRobotStatus.xBusy
			AND NOT stMagazineStatus.xBusy
			AND NOT xAnyMachineBusy
			AND NOT xMotionBusy;
		IF xReset AND xResetAllowed THEN
			Error.dwErrorLast := Error.dwErrorActive;
			Error.dwErrorActive := DWORD#0;
			IF NOT stRobotStatus.xBlankAvailable THEN
				uiBlankPayloadType := UINT#0;
			END_IF;
			IF NOT stRobotStatus.xDetailAvailable THEN
				uiDetailPayloadType := UINT#0;
			END_IF;
			eState := E_CELL_MANAGER_STATE.IDLE;
		END_IF;

	E_CELL_MANAGER_STATE.TEST_ABORT_STOP:
		xStopRequested := TRUE;
		Command.stRobot.xStop := TRUE;
		Command.stMagazine.xStop := TRUE;
		FOR uiMachine := FIRST_MACHINE TO LAST_MACHINE DO
			Command.axMachineExecute[uiMachine] := FALSE;
		END_FOR;
		IF NOT stRobotStatus.xBusy
		AND NOT xMotionBusy
		AND NOT stMagazineStatus.xBusy THEN
			xRunning := FALSE;
			xStopRequested := FALSE;
			xMachineServiceStarted := FALSE;
			xReselectAfterRobotRelease := FALSE;
			uiSelectedMachine := UINT#0;
			uiSelectedType := UINT#0;
			eMachineOperation := E_MACHINE_OPERATION.NONE;
			eMagazineOperation := E_MAGAZINE_OPERATION.NONE;
			eState := E_CELL_MANAGER_STATE.IDLE;
		END_IF;
END_CASE;

// Назначение фиксируется уже при планировании, до следующего RunTwoPallet.
// После загрузки заготовки владелец остаётся до PUT; отсутствие xBlankAvailable
// само по себе не разрешает смену палеты или переназначение готовой детали.
IF (uiActiveMagazine >= UINT#1) AND (uiActiveMagazine <= UINT#2) THEN
	IF (eState = E_CELL_MANAGER_STATE.MAGAZINE_EXECUTE)
	AND ((eMagazineOperation = E_MAGAZINE_OPERATION.TAKE)
		OR (eMagazineOperation = E_MAGAZINE_OPERATION.CHANGE)) THEN
		uiReturnMagazine := uiActiveMagazine;
	ELSIF (uiReturnMagazine = UINT#0)
	AND (eMachineOperation = E_MACHINE_OPERATION.UNLOAD)
	AND (eState = E_CELL_MANAGER_STATE.ROUTE_TO_TARGET) THEN
		uiReturnMagazine := uiActiveMagazine;
	END_IF;
END_IF;

// LOAD пустого станка и доставка на ГК завершаются без PUT. Публикуем
// освобождение в ТОМ ЖЕ вызове, который завершил операцию: RunTwoPallet
// следующего скана должен увидеть окно до нового планирования UNLOAD.
IF NOT stRobotStatus.xBusy
AND NOT stRobotStatus.xBlankAvailable
AND NOT stRobotStatus.xDetailAvailable
AND ((eState = E_CELL_MANAGER_STATE.IDLE)
	OR (eState = E_CELL_MANAGER_STATE.PLAN_TARGET)
	OR (eState = E_CELL_MANAGER_STATE.SELECT_FALLBACK)
	OR (eState = E_CELL_MANAGER_STATE.WAIT_MAGAZINE)) THEN
	uiReturnMagazine := UINT#0;
END_IF;

// Фиксируем позу только после завершённой штатной остановки или нормального
// окончания цикла. Аварийный переход оставляет xSafetyHomeRequired активным.
IF xWasRunning
AND NOT xRunning
AND (eState = E_CELL_MANAGER_STATE.IDLE)
AND NOT xSafetyHomeRequired THEN
	lrStoppedPoseX := lrRobotActualX;
	lrStoppedPoseY := lrRobotActualY;
	lrStoppedPoseZ := lrRobotActualZ;
	xStoppedPoseValid := TRUE;
END_IF;
xWasRunning := xRunning;

IF eState <> E_CELL_MANAGER_STATE.ERROR THEN
	xResetAllowed := FALSE;
END_IF;

Status.xMagazineExchangeAllowed := NOT xStopRequested
	AND ((eState = E_CELL_MANAGER_STATE.IDLE) OR (eState = E_CELL_MANAGER_STATE.PLAN_TARGET)
		OR (eState = E_CELL_MANAGER_STATE.WAIT_TARGET) OR (eState = E_CELL_MANAGER_STATE.WAIT_MAGAZINE));
Status.xRunning := xRunning;
Status.xStopPending := xStopRequested AND xRunning;
Status.xBusy := xRunning
	AND (eState <> E_CELL_MANAGER_STATE.IDLE)
	AND (eState <> E_CELL_MANAGER_STATE.ERROR);
Status.xWaitingMachine := (eState = E_CELL_MANAGER_STATE.WAIT_TARGET)
	OR (eState = E_CELL_MANAGER_STATE.SELECT_FALLBACK);
Status.xWaitingMagazine := eState = E_CELL_MANAGER_STATE.WAIT_MAGAZINE;
Status.xError := eState = E_CELL_MANAGER_STATE.ERROR;
Status.xReadyToStart := xReadyToStart;
Status.xStartAllowed := xReadyToStart
	OR (xRunning
		AND xStopRequested
		AND NOT xManual
		AND (eState <> E_CELL_MANAGER_STATE.MACHINE_FAULT_STOP));
Status.xStopAllowed := xRunning AND NOT xStopRequested;
Status.xResetAllowed := xResetAllowed;
// Ручной режим нельзя включить поверх работающего автоматического цикла.
// xManual уже отфильтрован до вызова FB, но это же условие публикуется HMI.
Status.xManualAllowed := NOT xRunning OR xGlobalError;
// В общей аварии оператору оставляем только ручное восстановление.
Status.xAutomaticAllowed := NOT xGlobalError AND NOT xIoEmergencyStopActive;
Status.xDrivesReady := xDrivesReady;
Status.xRobotReady := xRobotReady;
Status.xMagazineReady := xMagazineReady;
Status.xSafetyHomeRequired := xSafetyHomeRequired;
Status.xRobotAtSafetyHome := xRobotAtSafetyHome;
Status.xStartCheckCellIdle := xStartCheckCellIdle;
Status.xStartCheckAutomaticMode := xStartCheckAutomaticMode;
Status.xStartCheckNoBlockingError := xStartCheckNoBlockingError;
Status.xStartCheckRobotInterfaceReady := xStartCheckRobotInterfaceReady;
Status.xStartCheckConfigurationValid := xStartCheckConfigurationValid;
Status.xStartCheckPointsConfigured := xStartCheckPointsConfigured;
Status.xStartCheckDrivesReady := xStartCheckDrivesReady;
Status.xStartCheckRobotReady := xStartCheckRobotReady;
Status.xStartCheckMagazineReady := xStartCheckMagazineReady;
Status.xStartCheckTaskAvailable := xStartCheckTaskAvailable;
Status.xStartCheckSafetyHome := xStartCheckSafetyHome;
Status.xStartCheckSafety := xStartCheckSafety;
Status.uiStartConditionsMet := uiStartConditionsMet;
Status.uiStartConditionsTotal := UINT#12;
Status.uiReadyMachines := uiReadyMachines;
Status.uiSelectedMachine := uiSelectedMachine;
Status.uiActiveMagazine := uiActiveMagazine;
Status.eMagazineOperation := eMagazineOperation;
CASE eState OF
	E_CELL_MANAGER_STATE.WAIT_GRIPPER1_CONTENT: uiOperatorPrompt := UINT#1;
	E_CELL_MANAGER_STATE.WAIT_GRIPPER1_TYPE: uiOperatorPrompt := UINT#2;
	E_CELL_MANAGER_STATE.WAIT_GRIPPER2_CONTENT: uiOperatorPrompt := UINT#3;
	E_CELL_MANAGER_STATE.WAIT_GRIPPER2_TYPE: uiOperatorPrompt := UINT#4;
	E_CELL_MANAGER_STATE.WAIT_START_MACHINE: uiOperatorPrompt := UINT#5;
ELSE
	uiOperatorPrompt := UINT#0;
END_CASE;
Status.xOperatorPromptActive := uiOperatorPrompt <> UINT#0;
Status.xOperatorChoiceAllowed := Status.xOperatorPromptActive
	AND NOT xManual
	AND NOT xGlobalError
	AND (Error.dwErrorActive = DWORD#0)
	AND xRobotInterfaceReady
	AND xConfigurationValid
	AND xPointsConfigured
	AND xDrivesReady
	AND xRobotReady
	AND xMagazineReady
	AND (NOT xSafetyHomeRequired OR xRobotAtSafetyHome);
Status.xOperatorCancelAllowed := Status.xOperatorPromptActive;
Status.uiOperatorPrompt := uiOperatorPrompt;
Status.uiOperatorTypeMask := uiOperatorTypeMask;
Status.uiOperatorMachineMask := uiOperatorMachineMask;

// Во время TAKE/CHANGE тип будущей заготовки уже известен. Передаём его
// FB_ROBOT до закрытия первого захвата, чтобы авария между CLAMP и DONE не
// оставила физически взятую заготовку с типом 0.
IF ((eMagazineOperation = E_MAGAZINE_OPERATION.TAKE)
	OR (eMagazineOperation = E_MAGAZINE_OPERATION.CHANGE))
AND (uiSelectedType >= UINT#1)
AND (uiSelectedType <= Config.uiTypeCount) THEN
	Command.uiBlankPayloadType := uiSelectedType;
ELSE
	Command.uiBlankPayloadType := uiBlankPayloadType;
END_IF;
Command.uiDetailPayloadType := uiDetailPayloadType;

CASE eState OF
	E_CELL_MANAGER_STATE.IDLE: Diag.eState := E_CELL_STATE.IDLE;
	E_CELL_MANAGER_STATE.PRESTART_IDENTIFY,
	E_CELL_MANAGER_STATE.WAIT_GRIPPER1_CONTENT,
	E_CELL_MANAGER_STATE.WAIT_GRIPPER1_TYPE,
	E_CELL_MANAGER_STATE.WAIT_GRIPPER2_CONTENT,
	E_CELL_MANAGER_STATE.WAIT_GRIPPER2_TYPE,
	E_CELL_MANAGER_STATE.WAIT_START_MACHINE: Diag.eState := E_CELL_STATE.ROUTE_PAYLOAD;
	E_CELL_MANAGER_STATE.PLAN_TARGET, E_CELL_MANAGER_STATE.SELECT_FALLBACK: Diag.eState := E_CELL_STATE.SELECT_MACHINE;
	E_CELL_MANAGER_STATE.MAGAZINE_EXECUTE: Diag.eState := E_CELL_STATE.MAGAZINE;
	E_CELL_MANAGER_STATE.RELEASE_MAGAZINE: Diag.eState := E_CELL_STATE.RELEASE_MAGAZINE;
	E_CELL_MANAGER_STATE.ROUTE_TO_TARGET: Diag.eState := E_CELL_STATE.MOVE_TO_MACHINE;
	E_CELL_MANAGER_STATE.RELEASE_ROBOT_COMMAND: Diag.eState := E_CELL_STATE.RELEASE_ROBOT_COMMAND;
	E_CELL_MANAGER_STATE.WAIT_TARGET: Diag.eState := E_CELL_STATE.WAIT_MACHINE;
	E_CELL_MANAGER_STATE.SERVICE_TARGET: Diag.eState := E_CELL_STATE.SERVICE_MACHINE;
	E_CELL_MANAGER_STATE.MACHINE_FAULT_STOP: Diag.eState := E_CELL_STATE.SERVICE_MACHINE;
	E_CELL_MANAGER_STATE.WAIT_MAGAZINE: Diag.eState := E_CELL_STATE.WAIT_MAGAZINE;
	E_CELL_MANAGER_STATE.GEOMETRY_WAIT_FREE: Diag.eState := E_CELL_STATE.GEOMETRY_WAIT;
	E_CELL_MANAGER_STATE.GEOMETRY_DELIVER, E_CELL_MANAGER_STATE.GEOMETRY_RELEASE_COMMAND: Diag.eState := E_CELL_STATE.GEOMETRY_TRANSFER;
	E_CELL_MANAGER_STATE.TEST_ABORT_STOP: Diag.eState := E_CELL_STATE.IDLE;
	E_CELL_MANAGER_STATE.ERROR: Diag.eState := E_CELL_STATE.ERROR;
END_CASE;

CycleStatus.eState := eState;
CycleStatus.uiSelectedMachine := uiSelectedMachine;
CycleStatus.uiSelectedType := uiSelectedType;
CycleStatus.uiBlankPayloadType := uiBlankPayloadType;
CycleStatus.uiDetailPayloadType := uiDetailPayloadType;
CycleStatus.iTakeSlot := iTakeSlot;
CycleStatus.iPutSlot := iPutSlot;
CycleStatus.xReturningBlank := (eMagazineOperation = E_MAGAZINE_OPERATION.RETURN_BLANK)
	AND ((eState = E_CELL_MANAGER_STATE.MAGAZINE_EXECUTE)
		OR (eState = E_CELL_MANAGER_STATE.RELEASE_MAGAZINE));
CycleStatus.axMachineStartPending := axMachineStartPending;
CycleStatus.auiBlankCount := stMagazineStatus.stTypeStatus.auiBlankCount;
CycleStatus.auiDetailCount := stMagazineStatus.stTypeStatus.auiDetailCount;
CycleStatus.auiFreeCount := stMagazineStatus.stTypeStatus.auiFreeCount;

Error.dwAlarmActive := Error.dwErrorActive;
IF Error.dwErrorActive <> DWORD#0 THEN
	Error.dwErrorLast := Error.dwErrorActive;
END_IF;
Error.stErrorActive := UpdateErrorView(dwError := Error.dwErrorActive);
Error.stErrorLast := UpdateErrorView(dwError := Error.dwErrorLast);
FaultStatus.xResetAllowed := Status.xResetAllowed AND NOT FaultStatus.xBusy;
